(* IEC 61131-3 sources: plc-st-coding-agent/progress/evidence/f14_v13_self_20261113/jobs/custom_deepseek-v4pro (part 3) *)

(* ---- public-hard-05.patch_base_03.st ---- *)
FUNCTION_BLOCK MechanicalArmControl
VAR_INPUT
    ManualMode : BOOL;
    SingleStepMode : BOOL;
    SingleCycleMode : BOOL;
    ContinuousMode : BOOL;
    EmergencyStop : BOOL;
    Start : BOOL;
    DownButton : BOOL;
    UpButton : BOOL;
    LeftButton : BOOL;
    RightButton : BOOL;
    GripButton : BOOL;
    ReleaseButton : BOOL;
    DownLimitSwitch : BOOL;
    UpLimitSwitch : BOOL;
    LeftLimitSwitch : BOOL;
    RightLimitSwitch : BOOL;
    GripLimitSwitch : BOOL;
    ReleaseLimitSwitch : BOOL;
END_VAR
VAR_OUTPUT
    MoveDown : BOOL;
    MoveUp : BOOL;
    MoveLeft : BOOL;
    MoveRight : BOOL;
    ActivateGrip : BOOL;
    ActivateRelease : BOOL;
END_VAR
VAR
    local_startR : R_TRIG;
    tmp_first_scan : BOOL := TRUE;
    tmp_start_pulse : BOOL;
    tmp_not_estop : BOOL;
    tmp_ss_step : INT := 0;
    tmp_ss_busy : BOOL := FALSE;
    tmp_auto_running : BOOL := FALSE;
    tmp_auto_step : INT := 0;
    tmp_cmd_step : INT := 0;
    tmp_cmd_active : BOOL := FALSE;
    tmp_limit_reached : BOOL := FALSE;
END_VAR

(* ENGINEERING_CONTRACT
   Outputs MoveDown/Up/Left/Right/ActivateGrip/ActivateRelease:
   - Activate: manual while button=1, not at axis limit, and no opposite button (PUB001,PUB020); auto while current step active.
   - Retain: none latching; auto sequence state retained until completion/estop.
   - Reset: EmergencyStop=FALSE forces all outputs off and resets auto/single-step state (PUB005).
   - Same-scan: on limit true, previous output off; auto cycle can start next output in same scan (PUB003,PUB004).
   - Manual opposite-direction conflict inhibits both (PUB001 + shared rule).
   - Single-step Start edge only when not busy; ignored during running action (PUB002).
   - Single-cycle/continuous Start edge only when not running; continuous wraps at left completion (PUB003,PUB004).
   - Steps 0..7 = down, grip, up, right, down, release, up, left.
   - Grip/Release completion via GripLimitSwitch/ReleaseLimitSwitch (PUB001,PUB002).
   - Unspecified: mode change outside selected branch aborts/pauses per branch.
*)

(* CONTRACT_RULES [] *)

MoveDown := FALSE;
MoveUp := FALSE;
MoveLeft := FALSE;
MoveRight := FALSE;
ActivateGrip := FALSE;
ActivateRelease := FALSE;

tmp_not_estop := EmergencyStop; (* TRUE means no emergency stop triggered *)

local_startR(CLK := Start);
tmp_start_pulse := local_startR.Q AND NOT tmp_first_scan;
tmp_first_scan := FALSE;

tmp_cmd_active := FALSE;
tmp_cmd_step := 0;

IF NOT tmp_not_estop THEN
    tmp_ss_step := 0;
    tmp_ss_busy := FALSE;
    tmp_auto_running := FALSE;
    tmp_auto_step := 0;
    RETURN;
END_IF;

IF ManualMode THEN
    IF DownButton AND NOT UpButton AND NOT DownLimitSwitch THEN
        MoveDown := TRUE;
    END_IF;
    IF UpButton AND NOT DownButton AND NOT UpLimitSwitch THEN
        MoveUp := TRUE;
    END_IF;
    IF LeftButton AND NOT RightButton AND NOT LeftLimitSwitch THEN
        MoveLeft := TRUE;
    END_IF;
    IF RightButton AND NOT LeftButton AND NOT RightLimitSwitch THEN
        MoveRight := TRUE;
    END_IF;
    IF GripButton AND NOT ReleaseButton AND NOT GripLimitSwitch THEN
        ActivateGrip := TRUE;
    END_IF;
    IF ReleaseButton AND NOT GripButton AND NOT ReleaseLimitSwitch THEN
        ActivateRelease := TRUE;
    END_IF;

ELSIF SingleStepMode THEN
    IF tmp_start_pulse AND NOT tmp_ss_busy THEN
        tmp_ss_busy := TRUE;
    END_IF;

    IF tmp_ss_busy THEN
        tmp_limit_reached := FALSE;
        CASE tmp_ss_step OF
            0: tmp_limit_reached := DownLimitSwitch;
            1: tmp_limit_reached := GripLimitSwitch;
            2: tmp_limit_reached := UpLimitSwitch;
            3: tmp_limit_reached := RightLimitSwitch;
            4: tmp_limit_reached := DownLimitSwitch;
            5: tmp_limit_reached := ReleaseLimitSwitch;
            6: tmp_limit_reached := UpLimitSwitch;
            7: tmp_limit_reached := LeftLimitSwitch;
        END_CASE;

        IF tmp_limit_reached THEN
            tmp_ss_busy := FALSE;
            tmp_ss_step := tmp_ss_step + 1;
            IF tmp_ss_step > 7 THEN
                tmp_ss_step := 0;
            END_IF;
        ELSE
            tmp_cmd_step := tmp_ss_step;
            tmp_cmd_active := TRUE;
        END_IF;
    END_IF;

ELSIF SingleCycleMode OR ContinuousMode THEN
    IF tmp_start_pulse AND NOT tmp_auto_running THEN
        tmp_auto_running := TRUE;
        tmp_auto_step := 0;
    END_IF;

    IF tmp_auto_running THEN
        tmp_limit_reached := FALSE;
        CASE tmp_auto_step OF
            0: tmp_limit_reached := DownLimitSwitch;
            1: tmp_limit_reached := GripLimitSwitch;
            2: tmp_limit_reached := UpLimitSwitch;
            3: tmp_limit_reached := RightLimitSwitch;
            4: tmp_limit_reached := DownLimitSwitch;
            5: tmp_limit_reached := ReleaseLimitSwitch;
            6: tmp_limit_reached := UpLimitSwitch;
            7: tmp_limit_reached := LeftLimitSwitch;
        END_CASE;

        IF tmp_limit_reached THEN
            IF tmp_auto_step = 7 THEN
                IF ContinuousMode THEN
                    tmp_auto_step := 0; (* start next cycle *)
                ELSE
                    tmp_auto_running := FALSE;
                    tmp_auto_step := 0;
                END_IF;
            ELSE
                tmp_auto_step := tmp_auto_step + 1;
            END_IF;
        END_IF;

        IF tmp_auto_running THEN
            tmp_cmd_step := tmp_auto_step;
            tmp_cmd_active := TRUE;
        END_IF;
    END_IF;
END_IF;

IF tmp_cmd_active THEN
    CASE tmp_cmd_step OF
        0: MoveDown := TRUE;
        1: ActivateGrip := TRUE;
        2: MoveUp := TRUE;
        3: MoveRight := TRUE;
        4: MoveDown := TRUE;
        5: ActivateRelease := TRUE;
        6: MoveUp := TRUE;
        7: MoveLeft := TRUE;
    END_CASE;
END_IF;

END_FUNCTION_BLOCK

(* ---- public-hard-05.raw_candidate_01.st ---- *)
FUNCTION_BLOCK MechanicalArmControl
VAR_INPUT
    ManualMode : BOOL;
    SingleStepMode : BOOL;
    SingleCycleMode : BOOL;
    ContinuousMode : BOOL;
    EmergencyStop : BOOL;
    Start : BOOL;
    DownButton : BOOL;
    UpButton : BOOL;
    LeftButton : BOOL;
    RightButton : BOOL;
    GripButton : BOOL;
    ReleaseButton : BOOL;
    DownLimitSwitch : BOOL;
    UpLimitSwitch : BOOL;
    LeftLimitSwitch : BOOL;
    RightLimitSwitch : BOOL;
    GripLimitSwitch : BOOL;
    ReleaseLimitSwitch : BOOL;
END_VAR
VAR_OUTPUT
    MoveDown : BOOL;
    MoveUp : BOOL;
    MoveLeft : BOOL;
    MoveRight : BOOL;
    ActivateGrip : BOOL;
    ActivateRelease : BOOL;
END_VAR
VAR
    local_startR : R_TRIG;
    tmp_start_pulse : BOOL;
    tmp_not_estop : BOOL;
    tmp_ss_step : INT := 0;
    tmp_ss_busy : BOOL := FALSE;
    tmp_auto_running : BOOL := FALSE;
    tmp_auto_step : INT := 0;
    tmp_cmd_step : INT := 0;
    tmp_cmd_active : BOOL := FALSE;
    tmp_limit_reached : BOOL := FALSE;
END_VAR

(* ENGINEERING_CONTRACT
   Outputs MoveDown/Up/Left/Right/ActivateGrip/ActivateRelease:
   - Activate: manual while button=1, not at axis limit, and no opposite button (PUB001,PUB020); auto while current step active.
   - Retain: none latching; auto sequence state retained until completion/estop.
   - Reset: EmergencyStop=FALSE forces all outputs off and resets auto/single-step state (PUB005).
   - Same-scan: on limit true, previous output off; auto cycle can start next output in same scan (PUB003,PUB004).
   - Manual opposite-direction conflict inhibits both (PUB001 + shared rule).
   - Single-step Start edge only when not busy; ignored during running action (PUB002).
   - Single-cycle/continuous Start edge only when not running; continuous wraps at left completion (PUB003,PUB004).
   - Steps 0..7 = down, grip, up, right, down, release, up, left.
   - Grip/Release completion via GripLimitSwitch/ReleaseLimitSwitch (PUB001,PUB002).
   - Unspecified: mode change outside selected branch aborts/pauses per branch.
*)

(* CONTRACT_RULES [] *)

MoveDown := FALSE;
MoveUp := FALSE;
MoveLeft := FALSE;
MoveRight := FALSE;
ActivateGrip := FALSE;
ActivateRelease := FALSE;

tmp_not_estop := EmergencyStop; (* TRUE means no emergency stop triggered *)

local_startR(CLK := Start);
tmp_start_pulse := local_startR.Q;

tmp_cmd_active := FALSE;
tmp_cmd_step := 0;

IF NOT tmp_not_estop THEN
    tmp_ss_step := 0;
    tmp_ss_busy := FALSE;
    tmp_auto_running := FALSE;
    tmp_auto_step := 0;
    RETURN;
END_IF;

IF ManualMode THEN
    IF DownButton AND NOT UpButton AND NOT DownLimitSwitch THEN
        MoveDown := TRUE;
    END_IF;
    IF UpButton AND NOT DownButton AND NOT UpLimitSwitch THEN
        MoveUp := TRUE;
    END_IF;
    IF LeftButton AND NOT RightButton AND NOT LeftLimitSwitch THEN
        MoveLeft := TRUE;
    END_IF;
    IF RightButton AND NOT LeftButton AND NOT RightLimitSwitch THEN
        MoveRight := TRUE;
    END_IF;
    IF GripButton AND NOT ReleaseButton AND NOT GripLimitSwitch THEN
        ActivateGrip := TRUE;
    END_IF;
    IF ReleaseButton AND NOT GripButton AND NOT ReleaseLimitSwitch THEN
        ActivateRelease := TRUE;
    END_IF;

ELSIF SingleStepMode THEN
    IF tmp_start_pulse AND NOT tmp_ss_busy THEN
        tmp_ss_busy := TRUE;
    END_IF;

    IF tmp_ss_busy THEN
        tmp_limit_reached := FALSE;
        CASE tmp_ss_step OF
            0: tmp_limit_reached := DownLimitSwitch;
            1: tmp_limit_reached := GripLimitSwitch;
            2: tmp_limit_reached := UpLimitSwitch;
            3: tmp_limit_reached := RightLimitSwitch;
            4: tmp_limit_reached := DownLimitSwitch;
            5: tmp_limit_reached := ReleaseLimitSwitch;
            6: tmp_limit_reached := UpLimitSwitch;
            7: tmp_limit_reached := LeftLimitSwitch;
        END_CASE;

        IF tmp_limit_reached THEN
            tmp_ss_busy := FALSE;
            tmp_ss_step := tmp_ss_step + 1;
            IF tmp_ss_step > 7 THEN
                tmp_ss_step := 0;
            END_IF;
        ELSE
            tmp_cmd_step := tmp_ss_step;
            tmp_cmd_active := TRUE;
        END_IF;
    END_IF;

ELSIF SingleCycleMode OR ContinuousMode THEN
    IF tmp_start_pulse AND NOT tmp_auto_running THEN
        tmp_auto_running := TRUE;
        tmp_auto_step := 0;
    END_IF;

    IF tmp_auto_running THEN
        tmp_limit_reached := FALSE;
        CASE tmp_auto_step OF
            0: tmp_limit_reached := DownLimitSwitch;
            1: tmp_limit_reached := GripLimitSwitch;
            2: tmp_limit_reached := UpLimitSwitch;
            3: tmp_limit_reached := RightLimitSwitch;
            4: tmp_limit_reached := DownLimitSwitch;
            5: tmp_limit_reached := ReleaseLimitSwitch;
            6: tmp_limit_reached := UpLimitSwitch;
            7: tmp_limit_reached := LeftLimitSwitch;
        END_CASE;

        IF tmp_limit_reached THEN
            IF tmp_auto_step = 7 THEN
                IF ContinuousMode THEN
                    tmp_auto_step := 0; (* start next cycle *)
                ELSE
                    tmp_auto_running := FALSE;
                    tmp_auto_step := 0;
                END_IF;
            ELSE
                tmp_auto_step := tmp_auto_step + 1;
            END_IF;
        END_IF;

        IF tmp_auto_running THEN
            tmp_cmd_step := tmp_auto_step;
            tmp_cmd_active := TRUE;
        END_IF;
    END_IF;
END_IF;

IF tmp_cmd_active THEN
    CASE tmp_cmd_step OF
        0: MoveDown := TRUE;
        1: ActivateGrip := TRUE;
        2: MoveUp := TRUE;
        3: MoveRight := TRUE;
        4: MoveDown := TRUE;
        5: ActivateRelease := TRUE;
        6: MoveUp := TRUE;
        7: MoveLeft := TRUE;
    END_CASE;
END_IF;

END_FUNCTION_BLOCK

(* ---- public-hard-05.raw_candidate_02.st ---- *)
FUNCTION_BLOCK MechanicalArmControl
VAR_INPUT
    ManualMode : BOOL;
    SingleStepMode : BOOL;
    SingleCycleMode : BOOL;
    ContinuousMode : BOOL;
    EmergencyStop : BOOL;
    Start : BOOL;
    DownButton : BOOL;
    UpButton : BOOL;
    LeftButton : BOOL;
    RightButton : BOOL;
    GripButton : BOOL;
    ReleaseButton : BOOL;
    DownLimitSwitch : BOOL;
    UpLimitSwitch : BOOL;
    LeftLimitSwitch : BOOL;
    RightLimitSwitch : BOOL;
    GripLimitSwitch : BOOL;
    ReleaseLimitSwitch : BOOL;
END_VAR
VAR_OUTPUT
    MoveDown : BOOL;
    MoveUp : BOOL;
    MoveLeft : BOOL;
    MoveRight : BOOL;
    ActivateGrip : BOOL;
    ActivateRelease : BOOL;
END_VAR
VAR
    local_startR : R_TRIG;
    tmp_first_scan : BOOL := TRUE;
    tmp_start_pulse : BOOL;
    tmp_not_estop : BOOL;
    tmp_ss_step : INT := 0;
    tmp_ss_busy : BOOL := FALSE;
    tmp_auto_running : BOOL := FALSE;
    tmp_auto_step : INT := 0;
    tmp_cmd_step : INT := 0;
    tmp_cmd_active : BOOL := FALSE;
    tmp_limit_reached : BOOL := FALSE;
END_VAR

(* ENGINEERING_CONTRACT
   Outputs MoveDown/Up/Left/Right/ActivateGrip/ActivateRelease:
   - Activate: manual while button=1, not at axis limit, and no opposite button (PUB001,PUB020); auto while current step active.
   - Retain: none latching; auto sequence state retained until completion/estop.
   - Reset: EmergencyStop=FALSE forces all outputs off and resets auto/single-step state (PUB005).
   - Same-scan: on limit true, previous output off; auto cycle can start next output in same scan (PUB003,PUB004).
   - Manual opposite-direction conflict inhibits both (PUB001 + shared rule).
   - Single-step Start edge only when not busy; ignored during running action (PUB002).
   - Single-cycle/continuous Start edge only when not running; continuous wraps at left completion (PUB003,PUB004).
   - Steps 0..7 = down, grip, up, right, down, release, up, left.
   - Grip/Release completion via GripLimitSwitch/ReleaseLimitSwitch (PUB001,PUB002).
   - Unspecified: mode change outside selected branch aborts/pauses per branch.
*)

(* CONTRACT_RULES [] *)

MoveDown := FALSE;
MoveUp := FALSE;
MoveLeft := FALSE;
MoveRight := FALSE;
ActivateGrip := FALSE;
ActivateRelease := FALSE;

tmp_not_estop := EmergencyStop; (* TRUE means no emergency stop triggered *)

local_startR(CLK := Start);
tmp_start_pulse := local_startR.Q AND NOT tmp_first_scan;
tmp_first_scan := FALSE;

tmp_cmd_active := FALSE;
tmp_cmd_step := 0;

IF NOT tmp_not_estop THEN
    tmp_ss_step := 0;
    tmp_ss_busy := FALSE;
    tmp_auto_running := FALSE;
    tmp_auto_step := 0;
    RETURN;
END_IF;

IF ManualMode THEN
    IF DownButton AND NOT UpButton AND NOT DownLimitSwitch THEN
        MoveDown := TRUE;
    END_IF;
    IF UpButton AND NOT DownButton AND NOT UpLimitSwitch THEN
        MoveUp := TRUE;
    END_IF;
    IF LeftButton AND NOT RightButton AND NOT LeftLimitSwitch THEN
        MoveLeft := TRUE;
    END_IF;
    IF RightButton AND NOT LeftButton AND NOT RightLimitSwitch THEN
        MoveRight := TRUE;
    END_IF;
    IF GripButton AND NOT ReleaseButton AND NOT GripLimitSwitch THEN
        ActivateGrip := TRUE;
    END_IF;
    IF ReleaseButton AND NOT GripButton AND NOT ReleaseLimitSwitch THEN
        ActivateRelease := TRUE;
    END_IF;

ELSIF SingleStepMode THEN
    IF tmp_start_pulse AND NOT tmp_ss_busy THEN
        tmp_ss_busy := TRUE;
    END_IF;

    IF tmp_ss_busy THEN
        tmp_limit_reached := FALSE;
        CASE tmp_ss_step OF
            0: tmp_limit_reached := DownLimitSwitch;
            1: tmp_limit_reached := GripLimitSwitch;
            2: tmp_limit_reached := UpLimitSwitch;
            3: tmp_limit_reached := RightLimitSwitch;
            4: tmp_limit_reached := DownLimitSwitch;
            5: tmp_limit_reached := ReleaseLimitSwitch;
            6: tmp_limit_reached := UpLimitSwitch;
            7: tmp_limit_reached := LeftLimitSwitch;
        END_CASE;

        IF tmp_limit_reached THEN
            tmp_ss_busy := FALSE;
            tmp_ss_step := tmp_ss_step + 1;
            IF tmp_ss_step > 7 THEN
                tmp_ss_step := 0;
            END_IF;
        ELSE
            tmp_cmd_step := tmp_ss_step;
            tmp_cmd_active := TRUE;
        END_IF;
    END_IF;

ELSIF SingleCycleMode OR ContinuousMode THEN
    IF tmp_start_pulse AND NOT tmp_auto_running THEN
        tmp_auto_running := TRUE;
        tmp_auto_step := 0;
    END_IF;

    IF tmp_auto_running THEN
        tmp_limit_reached := FALSE;
        CASE tmp_auto_step OF
            0: tmp_limit_reached := DownLimitSwitch;
            1: tmp_limit_reached := GripLimitSwitch;
            2: tmp_limit_reached := UpLimitSwitch;
            3: tmp_limit_reached := RightLimitSwitch;
            4: tmp_limit_reached := DownLimitSwitch;
            5: tmp_limit_reached := ReleaseLimitSwitch;
            6: tmp_limit_reached := UpLimitSwitch;
            7: tmp_limit_reached := LeftLimitSwitch;
        END_CASE;

        IF tmp_limit_reached THEN
            IF tmp_auto_step = 7 THEN
                IF ContinuousMode THEN
                    tmp_auto_step := 0; (* start next cycle *)
                ELSE
                    tmp_auto_running := FALSE;
                    tmp_auto_step := 0;
                END_IF;
            ELSE
                tmp_auto_step := tmp_auto_step + 1;
            END_IF;
        END_IF;

        IF tmp_auto_running THEN
            tmp_cmd_step := tmp_auto_step;
            tmp_cmd_active := TRUE;
        END_IF;
    END_IF;
END_IF;

IF tmp_cmd_active THEN
    CASE tmp_cmd_step OF
        0: MoveDown := TRUE;
        1: ActivateGrip := TRUE;
        2: MoveUp := TRUE;
        3: MoveRight := TRUE;
        4: MoveDown := TRUE;
        5: ActivateRelease := TRUE;
        6: MoveUp := TRUE;
        7: MoveLeft := TRUE;
    END_CASE;
END_IF;

END_FUNCTION_BLOCK

(* ---- public-hard-05.raw_candidate_03.st ---- *)
FUNCTION_BLOCK MechanicalArmControl
VAR_INPUT
    ManualMode : BOOL;
    SingleStepMode : BOOL;
    SingleCycleMode : BOOL;
    ContinuousMode : BOOL;
    EmergencyStop : BOOL;
    Start : BOOL;
    DownButton : BOOL;
    UpButton : BOOL;
    LeftButton : BOOL;
    RightButton : BOOL;
    GripButton : BOOL;
    ReleaseButton : BOOL;
    DownLimitSwitch : BOOL;
    UpLimitSwitch : BOOL;
    LeftLimitSwitch : BOOL;
    RightLimitSwitch : BOOL;
    GripLimitSwitch : BOOL;
    ReleaseLimitSwitch : BOOL;
END_VAR
VAR_OUTPUT
    MoveDown : BOOL;
    MoveUp : BOOL;
    MoveLeft : BOOL;
    MoveRight : BOOL;
    ActivateGrip : BOOL;
    ActivateRelease : BOOL;
END_VAR
VAR
    local_startR : R_TRIG;
    tmp_start_pulse : BOOL;
    tmp_not_estop : BOOL;
    tmp_ss_step : INT := 0;
    tmp_ss_busy : BOOL := FALSE;
    tmp_auto_running : BOOL := FALSE;
    tmp_auto_step : INT := 0;
    tmp_cmd_step : INT := 0;
    tmp_cmd_active : BOOL := FALSE;
    tmp_limit_reached : BOOL := FALSE;
END_VAR

(* ENGINEERING_CONTRACT
   Outputs MoveDown/Up/Left/Right/ActivateGrip/ActivateRelease:
   - Activate: manual while button=1, not at axis limit, and no opposite button (PUB001,PUB020); auto while current step active.
   - Retain: none latching; auto sequence state retained until completion/estop.
   - Reset: EmergencyStop=FALSE forces all outputs off and resets auto/single-step state (PUB005).
   - Same-scan: on limit true, previous output off; auto cycle can start next output in same scan (PUB003,PUB004).
   - Manual opposite-direction conflict inhibits both (PUB001 + shared rule).
   - Single-step Start edge only when not busy; ignored during running action (PUB002).
   - Single-cycle/continuous Start edge only when not running; continuous wraps at left completion (PUB003,PUB004).
   - Steps 0..7 = down, grip, up, right, down, release, up, left.
   - Grip/Release completion via GripLimitSwitch/ReleaseLimitSwitch (PUB001,PUB002).
   - Unspecified: mode change outside selected branch aborts/pauses per branch.
*)

(* CONTRACT_RULES [] *)

MoveDown := FALSE;
MoveUp := FALSE;
MoveLeft := FALSE;
MoveRight := FALSE;
ActivateGrip := FALSE;
ActivateRelease := FALSE;

tmp_not_estop := EmergencyStop; (* TRUE means no emergency stop triggered *)

local_startR(CLK := Start);
tmp_start_pulse := local_startR.Q;

tmp_cmd_active := FALSE;
tmp_cmd_step := 0;

IF NOT tmp_not_estop THEN
    tmp_ss_step := 0;
    tmp_ss_busy := FALSE;
    tmp_auto_running := FALSE;
    tmp_auto_step := 0;
    RETURN;
END_IF;

IF ManualMode THEN
    IF DownButton AND NOT UpButton AND NOT DownLimitSwitch THEN
        MoveDown := TRUE;
    END_IF;
    IF UpButton AND NOT DownButton AND NOT UpLimitSwitch THEN
        MoveUp := TRUE;
    END_IF;
    IF LeftButton AND NOT RightButton AND NOT LeftLimitSwitch THEN
        MoveLeft := TRUE;
    END_IF;
    IF RightButton AND NOT LeftButton AND NOT RightLimitSwitch THEN
        MoveRight := TRUE;
    END_IF;
    IF GripButton AND NOT ReleaseButton AND NOT GripLimitSwitch THEN
        ActivateGrip := TRUE;
    END_IF;
    IF ReleaseButton AND NOT GripButton AND NOT ReleaseLimitSwitch THEN
        ActivateRelease := TRUE;
    END_IF;

ELSIF SingleStepMode THEN
    IF tmp_start_pulse AND NOT tmp_ss_busy THEN
        tmp_ss_busy := TRUE;
    END_IF;

    IF tmp_ss_busy THEN
        tmp_limit_reached := FALSE;
        CASE tmp_ss_step OF
            0: tmp_limit_reached := DownLimitSwitch;
            1: tmp_limit_reached := GripLimitSwitch;
            2: tmp_limit_reached := UpLimitSwitch;
            3: tmp_limit_reached := RightLimitSwitch;
            4: tmp_limit_reached := DownLimitSwitch;
            5: tmp_limit_reached := ReleaseLimitSwitch;
            6: tmp_limit_reached := UpLimitSwitch;
            7: tmp_limit_reached := LeftLimitSwitch;
        END_CASE;

        IF tmp_limit_reached THEN
            tmp_ss_busy := FALSE;
            tmp_ss_step := tmp_ss_step + 1;
            IF tmp_ss_step > 7 THEN
                tmp_ss_step := 0;
            END_IF;
        ELSE
            tmp_cmd_step := tmp_ss_step;
            tmp_cmd_active := TRUE;
        END_IF;
    END_IF;

ELSIF SingleCycleMode OR ContinuousMode THEN
    IF tmp_start_pulse AND NOT tmp_auto_running THEN
        tmp_auto_running := TRUE;
        tmp_auto_step := 0;
    END_IF;

    IF tmp_auto_running THEN
        tmp_limit_reached := FALSE;
        CASE tmp_auto_step OF
            0: tmp_limit_reached := DownLimitSwitch;
            1: tmp_limit_reached := GripLimitSwitch;
            2: tmp_limit_reached := UpLimitSwitch;
            3: tmp_limit_reached := RightLimitSwitch;
            4: tmp_limit_reached := DownLimitSwitch;
            5: tmp_limit_reached := ReleaseLimitSwitch;
            6: tmp_limit_reached := UpLimitSwitch;
            7: tmp_limit_reached := LeftLimitSwitch;
        END_CASE;

        IF tmp_limit_reached THEN
            IF tmp_auto_step = 7 THEN
                IF ContinuousMode THEN
                    tmp_auto_step := 0; (* start next cycle *)
                ELSE
                    tmp_auto_running := FALSE;
                    tmp_auto_step := 0;
                END_IF;
            ELSE
                tmp_auto_step := tmp_auto_step + 1;
            END_IF;
        END_IF;

        IF tmp_auto_running THEN
            tmp_cmd_step := tmp_auto_step;
            tmp_cmd_active := TRUE;
        END_IF;
    END_IF;
END_IF;

IF tmp_cmd_active THEN
    CASE tmp_cmd_step OF
        0: MoveDown := TRUE;
        1: ActivateGrip := TRUE;
        2: MoveUp := TRUE;
        3: MoveRight := TRUE;
        4: MoveDown := TRUE;
        5: ActivateRelease := TRUE;
        6: MoveUp := TRUE;
        7: MoveLeft := TRUE;
    END_CASE;
END_IF;

END_FUNCTION_BLOCK

(* ---- public-hard-06.candidate_01.st ---- *)
FUNCTION_BLOCK ProductionControl
VAR_INPUT
    Mode : BOOL;
    ForwardButton : BOOL;
    ReverseButton : BOOL;
    SensorFeed : BOOL;
    SensorWash : BOOL;
    SensorWeight : BOOL;
    SensorFiring : BOOL;
    SensorOutput : BOOL;
    washComplete : BOOL;
    weightComplete : BOOL;
    weight : REAL;
    firingComplete : BOOL;
END_VAR
VAR_OUTPUT
    MotorForward : BOOL;
    MotorReverse : BOOL;
    kick : BOOL;
    CompletionLight : BOOL;
    firingTemp : REAL;
END_VAR
VAR
    AutoStep : INT := 0;
    AutoInit : BOOL := FALSE;
    lastFiringTemp : REAL := 0.0;
    rtWash : R_TRIG;
    rtWeight : R_TRIG;
    rtFiring : R_TRIG;
    washEdge : BOOL;
    weightEdge : BOOL;
    firingEdge : BOOL;
    tmp_unqualified : BOOL;
END_VAR

(*
ENGINEERING_CONTRACT
MotorForward: auto active in states 10/30/50/70; manual = ForwardButton AND NOT ReverseButton.
MotorReverse: manual only, interlocked with ForwardButton; both false if both buttons true.
kick: pulse on rising weightComplete when weight < 100 or weight > 200 (unqualified).
CompletionLight: combinational = SensorOutput while Mode=TRUE; off in manual.
firingTemp: stored on qualified weightComplete; formula 500 + (weight-100)*0.5, retained otherwise.
Units: weight REAL in same unit as thresholds; firingTemp REAL degrees; boundaries inclusive 100..200.
*)
(* CONTRACT_RULES [] *)

rtWash(CLK := washComplete);
rtWeight(CLK := weightComplete);
rtFiring(CLK := firingComplete);
washEdge := rtWash.Q;
weightEdge := rtWeight.Q;
firingEdge := rtFiring.Q;

IF NOT AutoInit THEN
    AutoInit := TRUE;
    IF SensorOutput THEN
        AutoStep := 80;
    ELSIF SensorFiring THEN
        AutoStep := 60;
    ELSIF SensorWeight THEN
        AutoStep := 40;
    ELSIF SensorWash THEN
        AutoStep := 20;
    ELSIF SensorFeed THEN
        AutoStep := 10;
    ELSE
        AutoStep := 0;
    END_IF;
END_IF;

IF NOT Mode THEN
    MotorForward := ForwardButton AND (NOT ReverseButton);
    MotorReverse := ReverseButton AND (NOT ForwardButton);
    kick := FALSE;
    CompletionLight := FALSE;
    firingTemp := lastFiringTemp;
    RETURN;
END_IF;

MotorForward := FALSE;
MotorReverse := FALSE;
kick := FALSE;
CompletionLight := FALSE;

CASE AutoStep OF
    0:
        IF SensorFeed THEN
            AutoStep := 10;
        END_IF;

    10:
        IF SensorWash THEN
            AutoStep := 20;
        END_IF;

    20:
        IF washEdge THEN
            AutoStep := 30;
        END_IF;

    30:
        IF SensorWeight THEN
            AutoStep := 40;
        END_IF;

    40:
        IF weightEdge THEN
            tmp_unqualified := (weight < 100.0) OR (weight > 200.0);
            IF tmp_unqualified THEN
                kick := TRUE;
                AutoStep := 0;
            ELSE
                lastFiringTemp := 500.0 + (weight - 100.0) * 0.5;
                AutoStep := 50;
            END_IF;
        END_IF;

    50:
        IF SensorFiring THEN
            AutoStep := 60;
        END_IF;

    60:
        IF firingEdge THEN
            AutoStep := 70;
        END_IF;

    70:
        IF SensorOutput THEN
            AutoStep := 80;
        END_IF;

    80:
        ;
END_CASE;

MotorForward := (AutoStep = 10) OR (AutoStep = 30) OR (AutoStep = 50) OR (AutoStep = 70);
MotorReverse := FALSE;
CompletionLight := SensorOutput;
firingTemp := lastFiringTemp;
END_FUNCTION_BLOCK

(* ---- public-hard-06.candidate_02.st ---- *)
FUNCTION_BLOCK ProductionControl
VAR_INPUT
    Mode : BOOL;
    ForwardButton : BOOL;
    ReverseButton : BOOL;
    SensorFeed : BOOL;
    SensorWash : BOOL;
    SensorWeight : BOOL;
    SensorFiring : BOOL;
    SensorOutput : BOOL;
    washComplete : BOOL;
    weightComplete : BOOL;
    weight : REAL;
    firingComplete : BOOL;
END_VAR
VAR_OUTPUT
    MotorForward : BOOL;
    MotorReverse : BOOL;
    kick : BOOL;
    CompletionLight : BOOL;
    firingTemp : REAL;
END_VAR
VAR
    AutoStep : INT := 0;
    AutoInit : BOOL := FALSE;
    lastFiringTemp : REAL := 0.0;
    rtWash : R_TRIG;
    rtWeight : R_TRIG;
    rtFiring : R_TRIG;
    washEdge : BOOL;
    weightEdge : BOOL;
    firingEdge : BOOL;
    tmp_unqualified : BOOL;
END_VAR

(*
ENGINEERING_CONTRACT
MotorForward: auto active in states 10/30/50/70; manual = ForwardButton AND NOT ReverseButton.
MotorReverse: manual only, interlocked with ForwardButton; both false if both buttons true.
kick: pulse on rising weightComplete when weight < 100 or weight > 200 (unqualified).
CompletionLight: combinational = SensorOutput while Mode=TRUE; off in manual.
firingTemp: stored on qualified weightComplete; formula 500 + (weight-100)*0.5, retained otherwise.
Units: weight REAL in same unit as thresholds; firingTemp REAL degrees; boundaries inclusive 100..200.
*)
(* CONTRACT_RULES [] *)

rtWash(CLK := washComplete);
rtWeight(CLK := weightComplete);
rtFiring(CLK := firingComplete);
washEdge := rtWash.Q;
weightEdge := rtWeight.Q;
firingEdge := rtFiring.Q;

IF NOT AutoInit THEN
    AutoInit := TRUE;
    IF SensorOutput THEN
        AutoStep := 80;
    ELSIF SensorFiring THEN
        AutoStep := 60;
    ELSIF SensorWeight THEN
        AutoStep := 40;
    ELSIF SensorWash THEN
        AutoStep := 20;
    ELSIF SensorFeed THEN
        AutoStep := 10;
    ELSE
        AutoStep := 0;
    END_IF;
END_IF;

IF NOT Mode THEN
    MotorForward := ForwardButton AND (NOT ReverseButton);
    MotorReverse := ReverseButton AND (NOT ForwardButton);
    kick := FALSE;
    CompletionLight := FALSE;
    firingTemp := lastFiringTemp;
    RETURN;
END_IF;

MotorForward := FALSE;
MotorReverse := FALSE;
kick := FALSE;
CompletionLight := FALSE;

CASE AutoStep OF
    0:
        IF SensorFeed THEN
            AutoStep := 10;
        END_IF;

    10:
        IF SensorWash THEN
            AutoStep := 20;
        END_IF;

    20:
        IF washEdge THEN
            AutoStep := 30;
        END_IF;

    30:
        IF SensorWeight THEN
            AutoStep := 40;
        END_IF;

    40:
        IF weightEdge THEN
            tmp_unqualified := (weight < 100.0) OR (weight > 200.0);
            IF tmp_unqualified THEN
                kick := TRUE;
                AutoStep := 0;
            ELSE
                lastFiringTemp := 500.0 + (weight - 100.0) * 0.5;
                AutoStep := 50;
            END_IF;
        END_IF;

    50:
        IF SensorFiring THEN
            AutoStep := 60;
        END_IF;

    60:
        IF firingEdge THEN
            AutoStep := 70;
        END_IF;

    70:
        IF SensorOutput THEN
            AutoStep := 80;
        END_IF;

    80:
        IF NOT SensorOutput THEN
            AutoStep := 0;
        END_IF;
END_CASE;

MotorForward := (AutoStep = 10) OR (AutoStep = 30) OR (AutoStep = 50) OR (AutoStep = 70);
MotorReverse := FALSE;
CompletionLight := SensorOutput;
firingTemp := lastFiringTemp;
END_FUNCTION_BLOCK

(* ---- public-hard-06.candidate_03.st ---- *)
FUNCTION_BLOCK ProductionControl
VAR_INPUT
    Mode : BOOL;
    ForwardButton : BOOL;
    ReverseButton : BOOL;
    SensorFeed : BOOL;
    SensorWash : BOOL;
    SensorWeight : BOOL;
    SensorFiring : BOOL;
    SensorOutput : BOOL;
    washComplete : BOOL;
    weightComplete : BOOL;
    weight : REAL;
    firingComplete : BOOL;
END_VAR
VAR_OUTPUT
    MotorForward : BOOL;
    MotorReverse : BOOL;
    kick : BOOL;
    CompletionLight : BOOL;
    firingTemp : REAL;
END_VAR
VAR
    AutoStep : INT := 0;
    AutoInit : BOOL := FALSE;
    lastFiringTemp : REAL := 0.0;
    rtWash : R_TRIG;
    rtWeight : R_TRIG;
    rtFiring : R_TRIG;
    washEdge : BOOL;
    weightEdge : BOOL;
    firingEdge : BOOL;
    rtMode : R_TRIG;
    ModeRise : BOOL;
    tmp_unqualified : BOOL;
END_VAR

(*
ENGINEERING_CONTRACT
MotorForward: auto active in states 10/30/50/70; manual = ForwardButton AND NOT ReverseButton.
MotorReverse: manual only, interlocked with ForwardButton; both false if both buttons true.
kick: pulse on rising weightComplete when weight < 100 or weight > 200 (unqualified).
CompletionLight: combinational = SensorOutput while Mode=TRUE; off in manual.
firingTemp: stored on qualified weightComplete; formula 500 + (weight-100)*0.5, retained otherwise.
Units: weight REAL in same unit as thresholds; firingTemp REAL degrees; boundaries inclusive 100..200.
*)
(* CONTRACT_RULES [] *)

rtMode(CLK := Mode);
ModeRise := rtMode.Q;
rtWash(CLK := washComplete);
rtWeight(CLK := weightComplete);
rtFiring(CLK := firingComplete);
washEdge := rtWash.Q;
weightEdge := rtWeight.Q;
firingEdge := rtFiring.Q;

IF (NOT AutoInit) OR ModeRise THEN
    AutoInit := TRUE;
    IF SensorOutput THEN
        AutoStep := 80;
    ELSIF SensorFiring THEN
        AutoStep := 60;
    ELSIF SensorWeight THEN
        AutoStep := 40;
    ELSIF SensorWash THEN
        AutoStep := 20;
    ELSIF SensorFeed THEN
        AutoStep := 10;
    ELSE
        AutoStep := 0;
    END_IF;
END_IF;

IF NOT Mode THEN
    MotorForward := ForwardButton AND (NOT ReverseButton);
    MotorReverse := ReverseButton AND (NOT ForwardButton);
    kick := FALSE;
    CompletionLight := FALSE;
    firingTemp := lastFiringTemp;
    RETURN;
END_IF;

MotorForward := FALSE;
MotorReverse := FALSE;
kick := FALSE;
CompletionLight := FALSE;

CASE AutoStep OF
    0:
        IF SensorFeed THEN
            AutoStep := 10;
        END_IF;

    10:
        IF SensorWash THEN
            AutoStep := 20;
        END_IF;

    20:
        IF washEdge THEN
            AutoStep := 30;
        END_IF;

    30:
        IF SensorWeight THEN
            AutoStep := 40;
        END_IF;

    40:
        IF weightEdge THEN
            tmp_unqualified := (weight < 100.0) OR (weight > 200.0);
            IF tmp_unqualified THEN
                kick := TRUE;
                AutoStep := 0;
            ELSE
                lastFiringTemp := 500.0 + (weight - 100.0) * 0.5;
                AutoStep := 50;
            END_IF;
        END_IF;

    50:
        IF SensorFiring THEN
            AutoStep := 60;
        END_IF;

    60:
        IF firingEdge THEN
            AutoStep := 70;
        END_IF;

    70:
        IF SensorOutput THEN
            AutoStep := 80;
        END_IF;

    80:
        IF NOT SensorOutput THEN
            AutoStep := 0;
        END_IF;
END_CASE;

MotorForward := (AutoStep = 10) OR (AutoStep = 30) OR (AutoStep = 50) OR (AutoStep = 70);
MotorReverse := FALSE;
CompletionLight := SensorOutput;
firingTemp := lastFiringTemp;
END_FUNCTION_BLOCK

(* ---- public-hard-06.candidate_04.st ---- *)
FUNCTION_BLOCK ProductionControl
VAR_INPUT
    Mode : BOOL;
    ForwardButton : BOOL;
    ReverseButton : BOOL;
    SensorFeed : BOOL;
    SensorWash : BOOL;
    SensorWeight : BOOL;
    SensorFiring : BOOL;
    SensorOutput : BOOL;
    washComplete : BOOL;
    weightComplete : BOOL;
    weight : REAL;
    firingComplete : BOOL;
END_VAR
VAR_OUTPUT
    MotorForward : BOOL;
    MotorReverse : BOOL;
    kick : BOOL;
    CompletionLight : BOOL;
    firingTemp : REAL;
END_VAR
VAR
    AutoStep : INT := 0;
    AutoInit : BOOL := FALSE;
    lastFiringTemp : REAL := 0.0;
    rtWash : R_TRIG;
    rtWeight : R_TRIG;
    rtFiring : R_TRIG;
    washEdge : BOOL;
    weightEdge : BOOL;
    firingEdge : BOOL;
    rtMode : R_TRIG;
    ModeRise : BOOL;
    tmp_unqualified : BOOL;
END_VAR

(*
ENGINEERING_CONTRACT
MotorForward: auto active in states 10/30/50/70; manual = ForwardButton AND NOT ReverseButton.
MotorReverse: manual only, interlocked with ForwardButton; both false if both buttons true.
kick: pulse on rising weightComplete when weight < 100 or weight > 200 (unqualified).
CompletionLight: combinational = SensorOutput while Mode=TRUE; off in manual.
firingTemp: stored on qualified weightComplete; formula 500 + (weight-100)*0.5, retained otherwise.
Units: weight REAL in same unit as thresholds; firingTemp REAL degrees; boundaries inclusive 100..200.
*)
(* CONTRACT_RULES [] *)

rtMode(CLK := Mode);
ModeRise := rtMode.Q;
rtWash(CLK := washComplete);
rtWeight(CLK := weightComplete);
rtFiring(CLK := firingComplete);
washEdge := rtWash.Q;
weightEdge := rtWeight.Q;
firingEdge := rtFiring.Q;

IF (NOT AutoInit) OR ModeRise THEN
    AutoInit := TRUE;
    IF SensorOutput THEN
        AutoStep := 80;
    ELSIF SensorFiring THEN
        AutoStep := 60;
    ELSIF SensorWeight THEN
        AutoStep := 40;
    ELSIF SensorWash THEN
        AutoStep := 20;
    ELSIF SensorFeed THEN
        AutoStep := 10;
    ELSE
        AutoStep := 0;
    END_IF;
END_IF;

IF NOT Mode THEN
    MotorForward := ForwardButton AND (NOT ReverseButton);
    MotorReverse := ReverseButton AND (NOT ForwardButton);
    kick := FALSE;
    CompletionLight := FALSE;
    firingTemp := lastFiringTemp;
    RETURN;
END_IF;

MotorForward := FALSE;
MotorReverse := FALSE;
kick := FALSE;
CompletionLight := FALSE;

CASE AutoStep OF
    0:
        IF SensorFeed THEN
            AutoStep := 10;
        END_IF;

    10:
        IF SensorWash THEN
            AutoStep := 20;
        END_IF;

    20:
        IF washComplete THEN
            AutoStep := 30;
        END_IF;

    30:
        IF SensorWeight THEN
            AutoStep := 40;
        END_IF;

    40:
        IF weightComplete THEN
            tmp_unqualified := (weight < 100.0) OR (weight > 200.0);
            IF tmp_unqualified THEN
                kick := TRUE;
                AutoStep := 0;
            ELSE
                lastFiringTemp := 500.0 + (weight - 100.0) * 0.5;
                AutoStep := 50;
            END_IF;
        END_IF;

    50:
        IF SensorFiring THEN
            AutoStep := 60;
        END_IF;

    60:
        IF firingComplete THEN
            AutoStep := 70;
        END_IF;

    70:
        IF SensorOutput THEN
            AutoStep := 80;
        END_IF;

    80:
        IF NOT SensorOutput THEN
            AutoStep := 0;
        END_IF;
END_CASE;

MotorForward := (AutoStep = 10) OR (AutoStep = 30) OR (AutoStep = 50) OR (AutoStep = 70);
MotorReverse := FALSE;
CompletionLight := SensorOutput;
firingTemp := lastFiringTemp;
END_FUNCTION_BLOCK

(* ---- public-hard-06.patch_base_02.st ---- *)
FUNCTION_BLOCK ProductionControl
VAR_INPUT
    Mode : BOOL;
    ForwardButton : BOOL;
    ReverseButton : BOOL;
    SensorFeed : BOOL;
    SensorWash : BOOL;
    SensorWeight : BOOL;
    SensorFiring : BOOL;
    SensorOutput : BOOL;
    washComplete : BOOL;
    weightComplete : BOOL;
    weight : REAL;
    firingComplete : BOOL;
END_VAR
VAR_OUTPUT
    MotorForward : BOOL;
    MotorReverse : BOOL;
    kick : BOOL;
    CompletionLight : BOOL;
    firingTemp : REAL;
END_VAR
VAR
    AutoStep : INT := 0;
    AutoInit : BOOL := FALSE;
    lastFiringTemp : REAL := 0.0;
    rtWash : R_TRIG;
    rtWeight : R_TRIG;
    rtFiring : R_TRIG;
    washEdge : BOOL;
    weightEdge : BOOL;
    firingEdge : BOOL;
    tmp_unqualified : BOOL;
END_VAR

(*
ENGINEERING_CONTRACT
MotorForward: auto active in states 10/30/50/70; manual = ForwardButton AND NOT ReverseButton.
MotorReverse: manual only, interlocked with ForwardButton; both false if both buttons true.
kick: pulse on rising weightComplete when weight < 100 or weight > 200 (unqualified).
CompletionLight: combinational = SensorOutput while Mode=TRUE; off in manual.
firingTemp: stored on qualified weightComplete; formula 500 + (weight-100)*0.5, retained otherwise.
Units: weight REAL in same unit as thresholds; firingTemp REAL degrees; boundaries inclusive 100..200.
*)
(* CONTRACT_RULES [] *)

rtWash(CLK := washComplete);
rtWeight(CLK := weightComplete);
rtFiring(CLK := firingComplete);
washEdge := rtWash.Q;
weightEdge := rtWeight.Q;
firingEdge := rtFiring.Q;

IF NOT AutoInit THEN
    AutoInit := TRUE;
    IF SensorOutput THEN
        AutoStep := 80;
    ELSIF SensorFiring THEN
        AutoStep := 60;
    ELSIF SensorWeight THEN
        AutoStep := 40;
    ELSIF SensorWash THEN
        AutoStep := 20;
    ELSIF SensorFeed THEN
        AutoStep := 10;
    ELSE
        AutoStep := 0;
    END_IF;
END_IF;

IF NOT Mode THEN
    MotorForward := ForwardButton AND (NOT ReverseButton);
    MotorReverse := ReverseButton AND (NOT ForwardButton);
    kick := FALSE;
    CompletionLight := FALSE;
    firingTemp := lastFiringTemp;
    RETURN;
END_IF;

MotorForward := FALSE;
MotorReverse := FALSE;
kick := FALSE;
CompletionLight := FALSE;

CASE AutoStep OF
    0:
        IF SensorFeed THEN
            AutoStep := 10;
        END_IF;

    10:
        IF SensorWash THEN
            AutoStep := 20;
        END_IF;

    20:
        IF washEdge THEN
            AutoStep := 30;
        END_IF;

    30:
        IF SensorWeight THEN
            AutoStep := 40;
        END_IF;

    40:
        IF weightEdge THEN
            tmp_unqualified := (weight < 100.0) OR (weight > 200.0);
            IF tmp_unqualified THEN
                kick := TRUE;
                AutoStep := 0;
            ELSE
                lastFiringTemp := 500.0 + (weight - 100.0) * 0.5;
                AutoStep := 50;
            END_IF;
        END_IF;

    50:
        IF SensorFiring THEN
            AutoStep := 60;
        END_IF;

    60:
        IF firingEdge THEN
            AutoStep := 70;
        END_IF;

    70:
        IF SensorOutput THEN
            AutoStep := 80;
        END_IF;

    80:
        ;
END_CASE;

MotorForward := (AutoStep = 10) OR (AutoStep = 30) OR (AutoStep = 50) OR (AutoStep = 70);
MotorReverse := FALSE;
CompletionLight := SensorOutput;
firingTemp := lastFiringTemp;
END_FUNCTION_BLOCK

(* ---- public-hard-06.patch_base_03.st ---- *)
FUNCTION_BLOCK ProductionControl
VAR_INPUT
    Mode : BOOL;
    ForwardButton : BOOL;
    ReverseButton : BOOL;
    SensorFeed : BOOL;
    SensorWash : BOOL;
    SensorWeight : BOOL;
    SensorFiring : BOOL;
    SensorOutput : BOOL;
    washComplete : BOOL;
    weightComplete : BOOL;
    weight : REAL;
    firingComplete : BOOL;
END_VAR
VAR_OUTPUT
    MotorForward : BOOL;
    MotorReverse : BOOL;
    kick : BOOL;
    CompletionLight : BOOL;
    firingTemp : REAL;
END_VAR
VAR
    AutoStep : INT := 0;
    AutoInit : BOOL := FALSE;
    lastFiringTemp : REAL := 0.0;
    rtWash : R_TRIG;
    rtWeight : R_TRIG;
    rtFiring : R_TRIG;
    washEdge : BOOL;
    weightEdge : BOOL;
    firingEdge : BOOL;
    tmp_unqualified : BOOL;
END_VAR

(*
ENGINEERING_CONTRACT
MotorForward: auto active in states 10/30/50/70; manual = ForwardButton AND NOT ReverseButton.
MotorReverse: manual only, interlocked with ForwardButton; both false if both buttons true.
kick: pulse on rising weightComplete when weight < 100 or weight > 200 (unqualified).
CompletionLight: combinational = SensorOutput while Mode=TRUE; off in manual.
firingTemp: stored on qualified weightComplete; formula 500 + (weight-100)*0.5, retained otherwise.
Units: weight REAL in same unit as thresholds; firingTemp REAL degrees; boundaries inclusive 100..200.
*)
(* CONTRACT_RULES [] *)

rtWash(CLK := washComplete);
rtWeight(CLK := weightComplete);
rtFiring(CLK := firingComplete);
washEdge := rtWash.Q;
weightEdge := rtWeight.Q;
firingEdge := rtFiring.Q;

IF NOT AutoInit THEN
    AutoInit := TRUE;
    IF SensorOutput THEN
        AutoStep := 80;
    ELSIF SensorFiring THEN
        AutoStep := 60;
    ELSIF SensorWeight THEN
        AutoStep := 40;
    ELSIF SensorWash THEN
        AutoStep := 20;
    ELSIF SensorFeed THEN
        AutoStep := 10;
    ELSE
        AutoStep := 0;
    END_IF;
END_IF;

IF NOT Mode THEN
    MotorForward := ForwardButton AND (NOT ReverseButton);
    MotorReverse := ReverseButton AND (NOT ForwardButton);
    kick := FALSE;
    CompletionLight := FALSE;
    firingTemp := lastFiringTemp;
    RETURN;
END_IF;

MotorForward := FALSE;
MotorReverse := FALSE;
kick := FALSE;
CompletionLight := FALSE;

CASE AutoStep OF
    0:
        IF SensorFeed THEN
            AutoStep := 10;
        END_IF;

    10:
        IF SensorWash THEN
            AutoStep := 20;
        END_IF;

    20:
        IF washEdge THEN
            AutoStep := 30;
        END_IF;

    30:
        IF SensorWeight THEN
            AutoStep := 40;
        END_IF;

    40:
        IF weightEdge THEN
            tmp_unqualified := (weight < 100.0) OR (weight > 200.0);
            IF tmp_unqualified THEN
                kick := TRUE;
                AutoStep := 0;
            ELSE
                lastFiringTemp := 500.0 + (weight - 100.0) * 0.5;
                AutoStep := 50;
            END_IF;
        END_IF;

    50:
        IF SensorFiring THEN
            AutoStep := 60;
        END_IF;

    60:
        IF firingEdge THEN
            AutoStep := 70;
        END_IF;

    70:
        IF SensorOutput THEN
            AutoStep := 80;
        END_IF;

    80:
        IF NOT SensorOutput THEN
            AutoStep := 0;
        END_IF;
END_CASE;

MotorForward := (AutoStep = 10) OR (AutoStep = 30) OR (AutoStep = 50) OR (AutoStep = 70);
MotorReverse := FALSE;
CompletionLight := SensorOutput;
firingTemp := lastFiringTemp;
END_FUNCTION_BLOCK

(* ---- public-hard-06.patch_base_04.st ---- *)
FUNCTION_BLOCK ProductionControl
VAR_INPUT
    Mode : BOOL;
    ForwardButton : BOOL;
    ReverseButton : BOOL;
    SensorFeed : BOOL;
    SensorWash : BOOL;
    SensorWeight : BOOL;
    SensorFiring : BOOL;
    SensorOutput : BOOL;
    washComplete : BOOL;
    weightComplete : BOOL;
    weight : REAL;
    firingComplete : BOOL;
END_VAR
VAR_OUTPUT
    MotorForward : BOOL;
    MotorReverse : BOOL;
    kick : BOOL;
    CompletionLight : BOOL;
    firingTemp : REAL;
END_VAR
VAR
    AutoStep : INT := 0;
    AutoInit : BOOL := FALSE;
    lastFiringTemp : REAL := 0.0;
    rtWash : R_TRIG;
    rtWeight : R_TRIG;
    rtFiring : R_TRIG;
    washEdge : BOOL;
    weightEdge : BOOL;
    firingEdge : BOOL;
    rtMode : R_TRIG;
    ModeRise : BOOL;
    tmp_unqualified : BOOL;
END_VAR

(*
ENGINEERING_CONTRACT
MotorForward: auto active in states 10/30/50/70; manual = ForwardButton AND NOT ReverseButton.
MotorReverse: manual only, interlocked with ForwardButton; both false if both buttons true.
kick: pulse on rising weightComplete when weight < 100 or weight > 200 (unqualified).
CompletionLight: combinational = SensorOutput while Mode=TRUE; off in manual.
firingTemp: stored on qualified weightComplete; formula 500 + (weight-100)*0.5, retained otherwise.
Units: weight REAL in same unit as thresholds; firingTemp REAL degrees; boundaries inclusive 100..200.
*)
(* CONTRACT_RULES [] *)

rtMode(CLK := Mode);
ModeRise := rtMode.Q;
rtWash(CLK := washComplete);
rtWeight(CLK := weightComplete);
rtFiring(CLK := firingComplete);
washEdge := rtWash.Q;
weightEdge := rtWeight.Q;
firingEdge := rtFiring.Q;

IF (NOT AutoInit) OR ModeRise THEN
    AutoInit := TRUE;
    IF SensorOutput THEN
        AutoStep := 80;
    ELSIF SensorFiring THEN
        AutoStep := 60;
    ELSIF SensorWeight THEN
        AutoStep := 40;
    ELSIF SensorWash THEN
        AutoStep := 20;
    ELSIF SensorFeed THEN
        AutoStep := 10;
    ELSE
        AutoStep := 0;
    END_IF;
END_IF;

IF NOT Mode THEN
    MotorForward := ForwardButton AND (NOT ReverseButton);
    MotorReverse := ReverseButton AND (NOT ForwardButton);
    kick := FALSE;
    CompletionLight := FALSE;
    firingTemp := lastFiringTemp;
    RETURN;
END_IF;

MotorForward := FALSE;
MotorReverse := FALSE;
kick := FALSE;
CompletionLight := FALSE;

CASE AutoStep OF
    0:
        IF SensorFeed THEN
            AutoStep := 10;
        END_IF;

    10:
        IF SensorWash THEN
            AutoStep := 20;
        END_IF;

    20:
        IF washEdge THEN
            AutoStep := 30;
        END_IF;

    30:
        IF SensorWeight THEN
            AutoStep := 40;
        END_IF;

    40:
        IF weightEdge THEN
            tmp_unqualified := (weight < 100.0) OR (weight > 200.0);
            IF tmp_unqualified THEN
                kick := TRUE;
                AutoStep := 0;
            ELSE
                lastFiringTemp := 500.0 + (weight - 100.0) * 0.5;
                AutoStep := 50;
            END_IF;
        END_IF;

    50:
        IF SensorFiring THEN
            AutoStep := 60;
        END_IF;

    60:
        IF firingEdge THEN
            AutoStep := 70;
        END_IF;

    70:
        IF SensorOutput THEN
            AutoStep := 80;
        END_IF;

    80:
        IF NOT SensorOutput THEN
            AutoStep := 0;
        END_IF;
END_CASE;

MotorForward := (AutoStep = 10) OR (AutoStep = 30) OR (AutoStep = 50) OR (AutoStep = 70);
MotorReverse := FALSE;
CompletionLight := SensorOutput;
firingTemp := lastFiringTemp;
END_FUNCTION_BLOCK

(* ---- public-hard-06.raw_candidate_01.st ---- *)
FUNCTION_BLOCK ProductionControl
VAR_INPUT
    Mode : BOOL;
    ForwardButton : BOOL;
    ReverseButton : BOOL;
    SensorFeed : BOOL;
    SensorWash : BOOL;
    SensorWeight : BOOL;
    SensorFiring : BOOL;
    SensorOutput : BOOL;
    washComplete : BOOL;
    weightComplete : BOOL;
    weight : REAL;
    firingComplete : BOOL;
END_VAR
VAR_OUTPUT
    MotorForward : BOOL;
    MotorReverse : BOOL;
    kick : BOOL;
    CompletionLight : BOOL;
    firingTemp : REAL;
END_VAR
VAR
    AutoStep : INT := 0;
    AutoInit : BOOL := FALSE;
    lastFiringTemp : REAL := 0.0;
    rtWash : R_TRIG;
    rtWeight : R_TRIG;
    rtFiring : R_TRIG;
    washEdge : BOOL;
    weightEdge : BOOL;
    firingEdge : BOOL;
    tmp_unqualified : BOOL;
END_VAR

(*
ENGINEERING_CONTRACT
MotorForward: auto active in states 10/30/50/70; manual = ForwardButton AND NOT ReverseButton.
MotorReverse: manual only, interlocked with ForwardButton; both false if both buttons true.
kick: pulse on rising weightComplete when weight < 100 or weight > 200 (unqualified).
CompletionLight: combinational = SensorOutput while Mode=TRUE; off in manual.
firingTemp: stored on qualified weightComplete; formula 500 + (weight-100)*0.5, retained otherwise.
Units: weight REAL in same unit as thresholds; firingTemp REAL degrees; boundaries inclusive 100..200.
*)
(* CONTRACT_RULES [] *)

rtWash(CLK := washComplete);
rtWeight(CLK := weightComplete);
rtFiring(CLK := firingComplete);
washEdge := rtWash.Q;
weightEdge := rtWeight.Q;
firingEdge := rtFiring.Q;

IF NOT AutoInit THEN
    AutoInit := TRUE;
    IF SensorOutput THEN
        AutoStep := 80;
    ELSIF SensorFiring THEN
        AutoStep := 60;
    ELSIF SensorWeight THEN
        AutoStep := 40;
    ELSIF SensorWash THEN
        AutoStep := 20;
    ELSIF SensorFeed THEN
        AutoStep := 10;
    ELSE
        AutoStep := 0;
    END_IF;
END_IF;

IF NOT Mode THEN
    MotorForward := ForwardButton AND (NOT ReverseButton);
    MotorReverse := ReverseButton AND (NOT ForwardButton);
    kick := FALSE;
    CompletionLight := FALSE;
    firingTemp := lastFiringTemp;
    RETURN;
END_IF;

MotorForward := FALSE;
MotorReverse := FALSE;
kick := FALSE;
CompletionLight := FALSE;

CASE AutoStep OF
    0:
        IF SensorFeed THEN
            AutoStep := 10;
        END_IF;

    10:
        IF SensorWash THEN
            AutoStep := 20;
        END_IF;

    20:
        IF washEdge THEN
            AutoStep := 30;
        END_IF;

    30:
        IF SensorWeight THEN
            AutoStep := 40;
        END_IF;

    40:
        IF weightEdge THEN
            tmp_unqualified := (weight < 100.0) OR (weight > 200.0);
            IF tmp_unqualified THEN
                kick := TRUE;
                AutoStep := 0;
            ELSE
                lastFiringTemp := 500.0 + (weight - 100.0) * 0.5;
                AutoStep := 50;
            END_IF;
        END_IF;

    50:
        IF SensorFiring THEN
            AutoStep := 60;
        END_IF;

    60:
        IF firingEdge THEN
            AutoStep := 70;
        END_IF;

    70:
        IF SensorOutput THEN
            AutoStep := 80;
        END_IF;

    80:
        ;
END_CASE;

MotorForward := (AutoStep = 10) OR (AutoStep = 30) OR (AutoStep = 50) OR (AutoStep = 70);
MotorReverse := FALSE;
CompletionLight := SensorOutput;
firingTemp := lastFiringTemp;
END_FUNCTION_BLOCK

(* ---- public-hard-06.raw_candidate_02.st ---- *)
FUNCTION_BLOCK ProductionControl
VAR_INPUT
    Mode : BOOL;
    ForwardButton : BOOL;
    ReverseButton : BOOL;
    SensorFeed : BOOL;
    SensorWash : BOOL;
    SensorWeight : BOOL;
    SensorFiring : BOOL;
    SensorOutput : BOOL;
    washComplete : BOOL;
    weightComplete : BOOL;
    weight : REAL;
    firingComplete : BOOL;
END_VAR
VAR_OUTPUT
    MotorForward : BOOL;
    MotorReverse : BOOL;
    kick : BOOL;
    CompletionLight : BOOL;
    firingTemp : REAL;
END_VAR
VAR
    AutoStep : INT := 0;
    AutoInit : BOOL := FALSE;
    lastFiringTemp : REAL := 0.0;
    rtWash : R_TRIG;
    rtWeight : R_TRIG;
    rtFiring : R_TRIG;
    washEdge : BOOL;
    weightEdge : BOOL;
    firingEdge : BOOL;
    tmp_unqualified : BOOL;
END_VAR

(*
ENGINEERING_CONTRACT
MotorForward: auto active in states 10/30/50/70; manual = ForwardButton AND NOT ReverseButton.
MotorReverse: manual only, interlocked with ForwardButton; both false if both buttons true.
kick: pulse on rising weightComplete when weight < 100 or weight > 200 (unqualified).
CompletionLight: combinational = SensorOutput while Mode=TRUE; off in manual.
firingTemp: stored on qualified weightComplete; formula 500 + (weight-100)*0.5, retained otherwise.
Units: weight REAL in same unit as thresholds; firingTemp REAL degrees; boundaries inclusive 100..200.
*)
(* CONTRACT_RULES [] *)

rtWash(CLK := washComplete);
rtWeight(CLK := weightComplete);
rtFiring(CLK := firingComplete);
washEdge := rtWash.Q;
weightEdge := rtWeight.Q;
firingEdge := rtFiring.Q;

IF NOT AutoInit THEN
    AutoInit := TRUE;
    IF SensorOutput THEN
        AutoStep := 80;
    ELSIF SensorFiring THEN
        AutoStep := 60;
    ELSIF SensorWeight THEN
        AutoStep := 40;
    ELSIF SensorWash THEN
        AutoStep := 20;
    ELSIF SensorFeed THEN
        AutoStep := 10;
    ELSE
        AutoStep := 0;
    END_IF;
END_IF;

IF NOT Mode THEN
    MotorForward := ForwardButton AND (NOT ReverseButton);
    MotorReverse := ReverseButton AND (NOT ForwardButton);
    kick := FALSE;
    CompletionLight := FALSE;
    firingTemp := lastFiringTemp;
    RETURN;
END_IF;

MotorForward := FALSE;
MotorReverse := FALSE;
kick := FALSE;
CompletionLight := FALSE;

CASE AutoStep OF
    0:
        IF SensorFeed THEN
            AutoStep := 10;
        END_IF;

    10:
        IF SensorWash THEN
            AutoStep := 20;
        END_IF;

    20:
        IF washEdge THEN
            AutoStep := 30;
        END_IF;

    30:
        IF SensorWeight THEN
            AutoStep := 40;
        END_IF;

    40:
        IF weightEdge THEN
            tmp_unqualified := (weight < 100.0) OR (weight > 200.0);
            IF tmp_unqualified THEN
                kick := TRUE;
                AutoStep := 0;
            ELSE
                lastFiringTemp := 500.0 + (weight - 100.0) * 0.5;
                AutoStep := 50;
            END_IF;
        END_IF;

    50:
        IF SensorFiring THEN
            AutoStep := 60;
        END_IF;

    60:
        IF firingEdge THEN
            AutoStep := 70;
        END_IF;

    70:
        IF SensorOutput THEN
            AutoStep := 80;
        END_IF;

    80:
        IF NOT SensorOutput THEN
            AutoStep := 0;
        END_IF;
END_CASE;

MotorForward := (AutoStep = 10) OR (AutoStep = 30) OR (AutoStep = 50) OR (AutoStep = 70);
MotorReverse := FALSE;
CompletionLight := SensorOutput;
firingTemp := lastFiringTemp;
END_FUNCTION_BLOCK

(* ---- public-hard-06.raw_candidate_03.st ---- *)
FUNCTION_BLOCK ProductionControl
VAR_INPUT
    Mode : BOOL;
    ForwardButton : BOOL;
    ReverseButton : BOOL;
    SensorFeed : BOOL;
    SensorWash : BOOL;
    SensorWeight : BOOL;
    SensorFiring : BOOL;
    SensorOutput : BOOL;
    washComplete : BOOL;
    weightComplete : BOOL;
    weight : REAL;
    firingComplete : BOOL;
END_VAR
VAR_OUTPUT
    MotorForward : BOOL;
    MotorReverse : BOOL;
    kick : BOOL;
    CompletionLight : BOOL;
    firingTemp : REAL;
END_VAR
VAR
    AutoStep : INT := 0;
    AutoInit : BOOL := FALSE;
    lastFiringTemp : REAL := 0.0;
    rtWash : R_TRIG;
    rtWeight : R_TRIG;
    rtFiring : R_TRIG;
    washEdge : BOOL;
    weightEdge : BOOL;
    firingEdge : BOOL;
    rtMode : R_TRIG;
    ModeRise : BOOL;
    tmp_unqualified : BOOL;
END_VAR

(*
ENGINEERING_CONTRACT
MotorForward: auto active in states 10/30/50/70; manual = ForwardButton AND NOT ReverseButton.
MotorReverse: manual only, interlocked with ForwardButton; both false if both buttons true.
kick: pulse on rising weightComplete when weight < 100 or weight > 200 (unqualified).
CompletionLight: combinational = SensorOutput while Mode=TRUE; off in manual.
firingTemp: stored on qualified weightComplete; formula 500 + (weight-100)*0.5, retained otherwise.
Units: weight REAL in same unit as thresholds; firingTemp REAL degrees; boundaries inclusive 100..200.
*)
(* CONTRACT_RULES [] *)

rtMode(CLK := Mode);
ModeRise := rtMode.Q;
rtWash(CLK := washComplete);
rtWeight(CLK := weightComplete);
rtFiring(CLK := firingComplete);
washEdge := rtWash.Q;
weightEdge := rtWeight.Q;
firingEdge := rtFiring.Q;

IF (NOT AutoInit) OR ModeRise THEN
    AutoInit := TRUE;
    IF SensorOutput THEN
        AutoStep := 80;
    ELSIF SensorFiring THEN
        AutoStep := 60;
    ELSIF SensorWeight THEN
        AutoStep := 40;
    ELSIF SensorWash THEN
        AutoStep := 20;
    ELSIF SensorFeed THEN
        AutoStep := 10;
    ELSE
        AutoStep := 0;
    END_IF;
END_IF;

IF NOT Mode THEN
    MotorForward := ForwardButton AND (NOT ReverseButton);
    MotorReverse := ReverseButton AND (NOT ForwardButton);
    kick := FALSE;
    CompletionLight := FALSE;
    firingTemp := lastFiringTemp;
    RETURN;
END_IF;

MotorForward := FALSE;
MotorReverse := FALSE;
kick := FALSE;
CompletionLight := FALSE;

CASE AutoStep OF
    0:
        IF SensorFeed THEN
            AutoStep := 10;
        END_IF;

    10:
        IF SensorWash THEN
            AutoStep := 20;
        END_IF;

    20:
        IF washEdge THEN
            AutoStep := 30;
        END_IF;

    30:
        IF SensorWeight THEN
            AutoStep := 40;
        END_IF;

    40:
        IF weightEdge THEN
            tmp_unqualified := (weight < 100.0) OR (weight > 200.0);
            IF tmp_unqualified THEN
                kick := TRUE;
                AutoStep := 0;
            ELSE
                lastFiringTemp := 500.0 + (weight - 100.0) * 0.5;
                AutoStep := 50;
            END_IF;
        END_IF;

    50:
        IF SensorFiring THEN
            AutoStep := 60;
        END_IF;

    60:
        IF firingEdge THEN
            AutoStep := 70;
        END_IF;

    70:
        IF SensorOutput THEN
            AutoStep := 80;
        END_IF;

    80:
        IF NOT SensorOutput THEN
            AutoStep := 0;
        END_IF;
END_CASE;

MotorForward := (AutoStep = 10) OR (AutoStep = 30) OR (AutoStep = 50) OR (AutoStep = 70);
MotorReverse := FALSE;
CompletionLight := SensorOutput;
firingTemp := lastFiringTemp;
END_FUNCTION_BLOCK

(* ---- public-hard-06.raw_candidate_04.st ---- *)
FUNCTION_BLOCK ProductionControl
VAR_INPUT
    Mode : BOOL;
    ForwardButton : BOOL;
    ReverseButton : BOOL;
    SensorFeed : BOOL;
    SensorWash : BOOL;
    SensorWeight : BOOL;
    SensorFiring : BOOL;
    SensorOutput : BOOL;
    washComplete : BOOL;
    weightComplete : BOOL;
    weight : REAL;
    firingComplete : BOOL;
END_VAR
VAR_OUTPUT
    MotorForward : BOOL;
    MotorReverse : BOOL;
    kick : BOOL;
    CompletionLight : BOOL;
    firingTemp : REAL;
END_VAR
VAR
    AutoStep : INT := 0;
    AutoInit : BOOL := FALSE;
    lastFiringTemp : REAL := 0.0;
    rtWash : R_TRIG;
    rtWeight : R_TRIG;
    rtFiring : R_TRIG;
    washEdge : BOOL;
    weightEdge : BOOL;
    firingEdge : BOOL;
    rtMode : R_TRIG;
    ModeRise : BOOL;
    tmp_unqualified : BOOL;
END_VAR

(*
ENGINEERING_CONTRACT
MotorForward: auto active in states 10/30/50/70; manual = ForwardButton AND NOT ReverseButton.
MotorReverse: manual only, interlocked with ForwardButton; both false if both buttons true.
kick: pulse on rising weightComplete when weight < 100 or weight > 200 (unqualified).
CompletionLight: combinational = SensorOutput while Mode=TRUE; off in manual.
firingTemp: stored on qualified weightComplete; formula 500 + (weight-100)*0.5, retained otherwise.
Units: weight REAL in same unit as thresholds; firingTemp REAL degrees; boundaries inclusive 100..200.
*)
(* CONTRACT_RULES [] *)

rtMode(CLK := Mode);
ModeRise := rtMode.Q;
rtWash(CLK := washComplete);
rtWeight(CLK := weightComplete);
rtFiring(CLK := firingComplete);
washEdge := rtWash.Q;
weightEdge := rtWeight.Q;
firingEdge := rtFiring.Q;

IF (NOT AutoInit) OR ModeRise THEN
    AutoInit := TRUE;
    IF SensorOutput THEN
        AutoStep := 80;
    ELSIF SensorFiring THEN
        AutoStep := 60;
    ELSIF SensorWeight THEN
        AutoStep := 40;
    ELSIF SensorWash THEN
        AutoStep := 20;
    ELSIF SensorFeed THEN
        AutoStep := 10;
    ELSE
        AutoStep := 0;
    END_IF;
END_IF;

IF NOT Mode THEN
    MotorForward := ForwardButton AND (NOT ReverseButton);
    MotorReverse := ReverseButton AND (NOT ForwardButton);
    kick := FALSE;
    CompletionLight := FALSE;
    firingTemp := lastFiringTemp;
    RETURN;
END_IF;

MotorForward := FALSE;
MotorReverse := FALSE;
kick := FALSE;
CompletionLight := FALSE;

CASE AutoStep OF
    0:
        IF SensorFeed THEN
            AutoStep := 10;
        END_IF;

    10:
        IF SensorWash THEN
            AutoStep := 20;
        END_IF;

    20:
        IF washComplete THEN
            AutoStep := 30;
        END_IF;

    30:
        IF SensorWeight THEN
            AutoStep := 40;
        END_IF;

    40:
        IF weightComplete THEN
            tmp_unqualified := (weight < 100.0) OR (weight > 200.0);
            IF tmp_unqualified THEN
                kick := TRUE;
                AutoStep := 0;
            ELSE
                lastFiringTemp := 500.0 + (weight - 100.0) * 0.5;
                AutoStep := 50;
            END_IF;
        END_IF;

    50:
        IF SensorFiring THEN
            AutoStep := 60;
        END_IF;

    60:
        IF firingComplete THEN
            AutoStep := 70;
        END_IF;

    70:
        IF SensorOutput THEN
            AutoStep := 80;
        END_IF;

    80:
        IF NOT SensorOutput THEN
            AutoStep := 0;
        END_IF;
END_CASE;

MotorForward := (AutoStep = 10) OR (AutoStep = 30) OR (AutoStep = 50) OR (AutoStep = 70);
MotorReverse := FALSE;
CompletionLight := SensorOutput;
firingTemp := lastFiringTemp;
END_FUNCTION_BLOCK

(* ---- public-medium-01.candidate_01.st ---- *)
TYPE ST_Pump :
STRUCT
    priority : INT;
    selection : BOOL;
    RunComd : BOOL;
END_STRUCT
END_TYPE;

FUNCTION_BLOCK MultiPumpSwitchingControl
VAR_INPUT
    mode : BOOL;
    start : BOOL;
    stop : BOOL;
END_VAR
VAR_IN_OUT
    pumpGroup : ARRAY[1..5] OF ST_Pump;
END_VAR
VAR
    running : BOOL := FALSE;
    tmp_startPrev : BOOL := FALSE;
    tmp_i : INT;
    tmp_j : INT;
    tmp_k : INT;
    tmp_order : ARRAY[1..5] OF INT;
    tmp_isTop : ARRAY[1..5] OF BOOL;
    tmp_prioLeft : INT;
    tmp_prioRight : INT;
END_VAR

(* ENGINEERING_CONTRACT
- Mode select: PUB001/PUB003. mode FALSE=manual, TRUE=auto; outputs follow current mode each scan.
- Running latch: rising edge of start (PUB002) sets running=TRUE; stop=TRUE (PUB004) resets running=FALSE.
- Same-scan priority: stop overrides start; stop and start tests use final same-scan input values.
- Manual RunComd (PUB001/PUB003): RunComd[i] = running AND pumpGroup[i].selection, i=1..5.
- Auto RunComd (PUB001/PUB002): top 3 priorities selected each scan; larger priority wins.
  Ties are unspecified; this block breaks ties by lower array index.
  RunComd[i] = running AND tmp_isTop[i].
- Running state is retained across mode changes until stop; no unstated mode-change reset.
- Units/boundaries: array indices 1..5, priority INT, RunComd BOOL.
*)
(* CONTRACT_RULES [] *)

IF stop THEN
    running := FALSE;
ELSIF (NOT tmp_startPrev) AND start THEN
    running := TRUE;
END_IF;

tmp_startPrev := start;

IF NOT mode THEN
    FOR tmp_i := 1 TO 5 DO
        pumpGroup[tmp_i].RunComd := running AND pumpGroup[tmp_i].selection;
    END_FOR;
ELSE
    FOR tmp_i := 1 TO 5 DO
        tmp_order[tmp_i] := tmp_i;
        tmp_isTop[tmp_i] := FALSE;
    END_FOR;

    FOR tmp_i := 1 TO 4 DO
        FOR tmp_j := tmp_i + 1 TO 5 DO
            tmp_prioRight := pumpGroup[tmp_order[tmp_j]].priority;
            tmp_prioLeft := pumpGroup[tmp_order[tmp_i]].priority;
            IF tmp_prioRight > tmp_prioLeft THEN
                tmp_k := tmp_order[tmp_i];
                tmp_order[tmp_i] := tmp_order[tmp_j];
                tmp_order[tmp_j] := tmp_k;
            END_IF;
        END_FOR;
    END_FOR;

    FOR tmp_i := 1 TO 3 DO
        tmp_isTop[tmp_order[tmp_i]] := TRUE;
    END_FOR;

    FOR tmp_i := 1 TO 5 DO
        pumpGroup[tmp_i].RunComd := running AND tmp_isTop[tmp_i];
    END_FOR;
END_IF;

END_FUNCTION_BLOCK

(* ---- public-medium-01.candidate_02.st ---- *)
TYPE ST_Pump :
STRUCT
    priority : INT;
    selection : BOOL;
    RunComd : BOOL;
END_STRUCT
END_TYPE;

FUNCTION_BLOCK MultiPumpSwitchingControl
VAR_INPUT
    mode : BOOL;
    start : BOOL;
    stop : BOOL;
END_VAR
VAR_IN_OUT
    pumpGroup : ARRAY[1..5] OF ST_Pump;
END_VAR
VAR
    running : BOOL := FALSE;
    tmp_i : INT;
    tmp_j : INT;
    tmp_k : INT;
    tmp_order : ARRAY[1..5] OF INT;
    tmp_isTop : ARRAY[1..5] OF BOOL;
    tmp_prioLeft : INT;
    tmp_prioRight : INT;
END_VAR

(* ENGINEERING_CONTRACT
- Mode select: PUB001/PUB003. mode FALSE=manual, TRUE=auto; outputs follow current mode each scan.
- Running latch: level-sensitive set/reset. stop=TRUE (PUB004) resets running=FALSE; otherwise start=TRUE (PUB002) sets running=TRUE. Once set, running remains TRUE until stop even if start goes FALSE.
- Same-scan priority: stop overrides start; stop and start tests use final same-scan input values.
- Manual RunComd (PUB001/PUB003): RunComd[i] = running AND pumpGroup[i].selection, i=1..5.
- Auto RunComd (PUB001/PUB002): top 3 priorities selected each scan; larger priority wins.
  Ties are unspecified; this block breaks ties by lower array index.
  RunComd[i] = running AND tmp_isTop[i].
- Running state is retained across mode changes until stop; no unstated mode-change reset.
- Units/boundaries: array indices 1..5, priority INT, RunComd BOOL.
*)
(* CONTRACT_RULES [] *)

IF stop THEN
    running := FALSE;
ELSIF start THEN
    running := TRUE;
END_IF;

IF NOT mode THEN
    FOR tmp_i := 1 TO 5 DO
        pumpGroup[tmp_i].RunComd := running AND pumpGroup[tmp_i].selection;
    END_FOR;
ELSE
    FOR tmp_i := 1 TO 5 DO
        tmp_order[tmp_i] := tmp_i;
        tmp_isTop[tmp_i] := FALSE;
    END_FOR;

    FOR tmp_i := 1 TO 4 DO
        FOR tmp_j := tmp_i + 1 TO 5 DO
            tmp_prioRight := pumpGroup[tmp_order[tmp_j]].priority;
            tmp_prioLeft := pumpGroup[tmp_order[tmp_i]].priority;
            IF tmp_prioRight > tmp_prioLeft THEN
                tmp_k := tmp_order[tmp_i];
                tmp_order[tmp_i] := tmp_order[tmp_j];
                tmp_order[tmp_j] := tmp_k;
            END_IF;
        END_FOR;
    END_FOR;

    FOR tmp_i := 1 TO 3 DO
        tmp_isTop[tmp_order[tmp_i]] := TRUE;
    END_FOR;

    FOR tmp_i := 1 TO 5 DO
        pumpGroup[tmp_i].RunComd := running AND tmp_isTop[tmp_i];
    END_FOR;
END_IF;

END_FUNCTION_BLOCK

(* ---- public-medium-01.patch_base_02.st ---- *)
TYPE ST_Pump :
STRUCT
    priority : INT;
    selection : BOOL;
    RunComd : BOOL;
END_STRUCT
END_TYPE;

FUNCTION_BLOCK MultiPumpSwitchingControl
VAR_INPUT
    mode : BOOL;
    start : BOOL;
    stop : BOOL;
END_VAR
VAR_IN_OUT
    pumpGroup : ARRAY[1..5] OF ST_Pump;
END_VAR
VAR
    running : BOOL := FALSE;
    tmp_startPrev : BOOL := FALSE;
    tmp_i : INT;
    tmp_j : INT;
    tmp_k : INT;
    tmp_order : ARRAY[1..5] OF INT;
    tmp_isTop : ARRAY[1..5] OF BOOL;
    tmp_prioLeft : INT;
    tmp_prioRight : INT;
END_VAR

(* ENGINEERING_CONTRACT
- Mode select: PUB001/PUB003. mode FALSE=manual, TRUE=auto; outputs follow current mode each scan.
- Running latch: rising edge of start (PUB002) sets running=TRUE; stop=TRUE (PUB004) resets running=FALSE.
- Same-scan priority: stop overrides start; stop and start tests use final same-scan input values.
- Manual RunComd (PUB001/PUB003): RunComd[i] = running AND pumpGroup[i].selection, i=1..5.
- Auto RunComd (PUB001/PUB002): top 3 priorities selected each scan; larger priority wins.
  Ties are unspecified; this block breaks ties by lower array index.
  RunComd[i] = running AND tmp_isTop[i].
- Running state is retained across mode changes until stop; no unstated mode-change reset.
- Units/boundaries: array indices 1..5, priority INT, RunComd BOOL.
*)
(* CONTRACT_RULES [] *)

IF stop THEN
    running := FALSE;
ELSIF (NOT tmp_startPrev) AND start THEN
    running := TRUE;
END_IF;

tmp_startPrev := start;

IF NOT mode THEN
    FOR tmp_i := 1 TO 5 DO
        pumpGroup[tmp_i].RunComd := running AND pumpGroup[tmp_i].selection;
    END_FOR;
ELSE
    FOR tmp_i := 1 TO 5 DO
        tmp_order[tmp_i] := tmp_i;
        tmp_isTop[tmp_i] := FALSE;
    END_FOR;

    FOR tmp_i := 1 TO 4 DO
        FOR tmp_j := tmp_i + 1 TO 5 DO
            tmp_prioRight := pumpGroup[tmp_order[tmp_j]].priority;
            tmp_prioLeft := pumpGroup[tmp_order[tmp_i]].priority;
            IF tmp_prioRight > tmp_prioLeft THEN
                tmp_k := tmp_order[tmp_i];
                tmp_order[tmp_i] := tmp_order[tmp_j];
                tmp_order[tmp_j] := tmp_k;
            END_IF;
        END_FOR;
    END_FOR;

    FOR tmp_i := 1 TO 3 DO
        tmp_isTop[tmp_order[tmp_i]] := TRUE;
    END_FOR;

    FOR tmp_i := 1 TO 5 DO
        pumpGroup[tmp_i].RunComd := running AND tmp_isTop[tmp_i];
    END_FOR;
END_IF;

END_FUNCTION_BLOCK

(* ---- public-medium-01.raw_candidate_01.st ---- *)
TYPE ST_Pump :
STRUCT
    priority : INT;
    selection : BOOL;
    RunComd : BOOL;
END_STRUCT
END_TYPE

FUNCTION_BLOCK MultiPumpSwitchingControl
VAR_INPUT
    mode : BOOL;
    start : BOOL;
    stop : BOOL;
END_VAR
VAR_IN_OUT
    pumpGroup : ARRAY[1..5] OF ST_Pump;
END_VAR
VAR
    running : BOOL := FALSE;
    tmp_startPrev : BOOL := FALSE;
    tmp_i : INT;
    tmp_j : INT;
    tmp_k : INT;
    tmp_order : ARRAY[1..5] OF INT;
    tmp_isTop : ARRAY[1..5] OF BOOL;
    tmp_prioLeft : INT;
    tmp_prioRight : INT;
END_VAR

(* ENGINEERING_CONTRACT
- Mode select: PUB001/PUB003. mode FALSE=manual, TRUE=auto; outputs follow current mode each scan.
- Running latch: rising edge of start (PUB002) sets running=TRUE; stop=TRUE (PUB004) resets running=FALSE.
- Same-scan priority: stop overrides start; stop and start tests use final same-scan input values.
- Manual RunComd (PUB001/PUB003): RunComd[i] = running AND pumpGroup[i].selection, i=1..5.
- Auto RunComd (PUB001/PUB002): top 3 priorities selected each scan; larger priority wins.
  Ties are unspecified; this block breaks ties by lower array index.
  RunComd[i] = running AND tmp_isTop[i].
- Running state is retained across mode changes until stop; no unstated mode-change reset.
- Units/boundaries: array indices 1..5, priority INT, RunComd BOOL.
*)
(* CONTRACT_RULES [] *)

IF stop THEN
    running := FALSE;
ELSIF (NOT tmp_startPrev) AND start THEN
    running := TRUE;
END_IF;

tmp_startPrev := start;

IF NOT mode THEN
    FOR tmp_i := 1 TO 5 DO
        pumpGroup[tmp_i].RunComd := running AND pumpGroup[tmp_i].selection;
    END_FOR;
ELSE
    FOR tmp_i := 1 TO 5 DO
        tmp_order[tmp_i] := tmp_i;
        tmp_isTop[tmp_i] := FALSE;
    END_FOR;

    FOR tmp_i := 1 TO 4 DO
        FOR tmp_j := tmp_i + 1 TO 5 DO
            tmp_prioRight := pumpGroup[tmp_order[tmp_j]].priority;
            tmp_prioLeft := pumpGroup[tmp_order[tmp_i]].priority;
            IF tmp_prioRight > tmp_prioLeft THEN
                tmp_k := tmp_order[tmp_i];
                tmp_order[tmp_i] := tmp_order[tmp_j];
                tmp_order[tmp_j] := tmp_k;
            END_IF;
        END_FOR;
    END_FOR;

    FOR tmp_i := 1 TO 3 DO
        tmp_isTop[tmp_order[tmp_i]] := TRUE;
    END_FOR;

    FOR tmp_i := 1 TO 5 DO
        pumpGroup[tmp_i].RunComd := running AND tmp_isTop[tmp_i];
    END_FOR;
END_IF;

END_FUNCTION_BLOCK

(* ---- public-medium-01.raw_candidate_02.st ---- *)
TYPE ST_Pump :
STRUCT
    priority : INT;
    selection : BOOL;
    RunComd : BOOL;
END_STRUCT
END_TYPE;

FUNCTION_BLOCK MultiPumpSwitchingControl
VAR_INPUT
    mode : BOOL;
    start : BOOL;
    stop : BOOL;
END_VAR
VAR_IN_OUT
    pumpGroup : ARRAY[1..5] OF ST_Pump;
END_VAR
VAR
    running : BOOL := FALSE;
    tmp_i : INT;
    tmp_j : INT;
    tmp_k : INT;
    tmp_order : ARRAY[1..5] OF INT;
    tmp_isTop : ARRAY[1..5] OF BOOL;
    tmp_prioLeft : INT;
    tmp_prioRight : INT;
END_VAR

(* ENGINEERING_CONTRACT
- Mode select: PUB001/PUB003. mode FALSE=manual, TRUE=auto; outputs follow current mode each scan.
- Running latch: level-sensitive set/reset. stop=TRUE (PUB004) resets running=FALSE; otherwise start=TRUE (PUB002) sets running=TRUE. Once set, running remains TRUE until stop even if start goes FALSE.
- Same-scan priority: stop overrides start; stop and start tests use final same-scan input values.
- Manual RunComd (PUB001/PUB003): RunComd[i] = running AND pumpGroup[i].selection, i=1..5.
- Auto RunComd (PUB001/PUB002): top 3 priorities selected each scan; larger priority wins.
  Ties are unspecified; this block breaks ties by lower array index.
  RunComd[i] = running AND tmp_isTop[i].
- Running state is retained across mode changes until stop; no unstated mode-change reset.
- Units/boundaries: array indices 1..5, priority INT, RunComd BOOL.
*)
(* CONTRACT_RULES [] *)

IF stop THEN
    running := FALSE;
ELSIF start THEN
    running := TRUE;
END_IF;

IF NOT mode THEN
    FOR tmp_i := 1 TO 5 DO
        pumpGroup[tmp_i].RunComd := running AND pumpGroup[tmp_i].selection;
    END_FOR;
ELSE
    FOR tmp_i := 1 TO 5 DO
        tmp_order[tmp_i] := tmp_i;
        tmp_isTop[tmp_i] := FALSE;
    END_FOR;

    FOR tmp_i := 1 TO 4 DO
        FOR tmp_j := tmp_i + 1 TO 5 DO
            tmp_prioRight := pumpGroup[tmp_order[tmp_j]].priority;
            tmp_prioLeft := pumpGroup[tmp_order[tmp_i]].priority;
            IF tmp_prioRight > tmp_prioLeft THEN
                tmp_k := tmp_order[tmp_i];
                tmp_order[tmp_i] := tmp_order[tmp_j];
                tmp_order[tmp_j] := tmp_k;
            END_IF;
        END_FOR;
    END_FOR;

    FOR tmp_i := 1 TO 3 DO
        tmp_isTop[tmp_order[tmp_i]] := TRUE;
    END_FOR;

    FOR tmp_i := 1 TO 5 DO
        pumpGroup[tmp_i].RunComd := running AND tmp_isTop[tmp_i];
    END_FOR;
END_IF;

END_FUNCTION_BLOCK

(* ---- public-medium-02.candidate_01.st ---- *)
TYPE ST_AnalogChannel :
STRUCT
    enable : BOOL;
    hiLIM : REAL;
    loLIM : REAL;
    bipolar : BOOL;
    measuringMode : INT;
    retVal : WORD;
    outputValue : REAL;
END_STRUCT
END_TYPE;

(* ENGINEERING_CONTRACT
   Loop count: count limited to 0..min(array lengths); ordinal start at each array lower bound (PUB001).
   channels[].retVal: activated on enabled scan; invalid mode -> 16#8001, invalid limits -> 16#8002,
   success -> 0 (PUB006, PUB007, PUB008).
   channels[].outputValue: written only on successful conversion; mode 0 linear scaling,
   mode 1 /10, mode 2 /100 (PUB003, PUB004, PUB005).
   Disabled channels retain prior retVal/outputValue (unspecified retention interpretation).
*)

(* CONTRACT_RULES [] *)

FUNCTION_BLOCK AnalogBatchProcessing
VAR_INPUT
    count : DINT;
END_VAR
VAR_IN_OUT
    analogValues : ARRAY[*] OF INT;
    channels : ARRAY[*] OF ST_AnalogChannel;
END_VAR
VAR
    local_i : DINT;
    local_n : DINT;
    local_analog_idx : DINT;
    local_channel_idx : DINT;
    local_raw : INT;
    local_mode : INT;
    local_min_len : DINT;
    local_ch_len : DINT;
    local_raw_min : REAL;
    local_raw_max : REAL;
    local_span_raw : REAL;
    local_ratio : REAL;
END_VAR

local_n := count;
IF local_n < 0 THEN
    local_n := 0;
END_IF;

local_min_len := UPPER_BOUND(analogValues, 1) - LOWER_BOUND(analogValues, 1) + 1;
local_ch_len := UPPER_BOUND(channels, 1) - LOWER_BOUND(channels, 1) + 1;
IF local_min_len > local_ch_len THEN
    local_min_len := local_ch_len;
END_IF;
IF local_n > local_min_len THEN
    local_n := local_min_len;
END_IF;

IF local_n > 0 THEN
    FOR local_i := 0 TO local_n - 1 DO
        local_analog_idx := LOWER_BOUND(analogValues, 1) + local_i;
        local_channel_idx := LOWER_BOUND(channels, 1) + local_i;

        IF channels[local_channel_idx].enable THEN
            local_mode := channels[local_channel_idx].measuringMode;

            IF (local_mode <> 0) AND (local_mode <> 1) AND (local_mode <> 2) THEN
                channels[local_channel_idx].retVal := 16#8001;
                (* skip conversion: outputValue unchanged *)
            ELSIF channels[local_channel_idx].hiLIM <= channels[local_channel_idx].loLIM THEN
                channels[local_channel_idx].retVal := 16#8002;
                (* skip conversion: outputValue unchanged *)
            ELSE
                channels[local_channel_idx].retVal := 0;
                CASE local_mode OF
                    0:
                        local_raw := analogValues[local_analog_idx];
                        IF channels[local_channel_idx].bipolar THEN
                            local_raw_min := -27648.0;
                            local_raw_max := 27648.0;
                        ELSE
                            local_raw_min := 0.0;
                            local_raw_max := 27648.0;
                        END_IF;

                        local_span_raw := local_raw_max - local_raw_min;
                        local_ratio := (TO_REAL(local_raw) - local_raw_min) / local_span_raw;
                        channels[local_channel_idx].outputValue := channels[local_channel_idx].loLIM
                            + local_ratio * (channels[local_channel_idx].hiLIM - channels[local_channel_idx].loLIM);

                    1:
                        channels[local_channel_idx].outputValue := TO_REAL(analogValues[local_analog_idx]) / 10.0;

                    2:
                        channels[local_channel_idx].outputValue := TO_REAL(analogValues[local_analog_idx]) / 100.0;
                END_CASE;
            END_IF;
        ELSE
            (* disabled: no writes to retVal or outputValue *)
        END_IF;
    END_FOR;
END_IF;

(* ---- public-medium-02.candidate_02.st ---- *)
TYPE ST_AnalogChannel :
STRUCT
    enable : BOOL;
    hiLIM : REAL;
    loLIM : REAL;
    bipolar : BOOL;
    measuringMode : INT;
    retVal : WORD;
    outputValue : REAL;
END_STRUCT
END_TYPE;

(* ENGINEERING_CONTRACT
   Loop count: count limited to 0..min(array lengths); ordinal start at each array lower bound (PUB001).
   channels[].retVal: activated on enabled scan; invalid mode -> 16#8001, invalid limits -> 16#8002,
   success -> 0 (PUB006, PUB007, PUB008).
   channels[].outputValue: written only on successful conversion; mode 0 linear scaling,
   mode 1 /10, mode 2 /100 (PUB003, PUB004, PUB005).
   Disabled channels retain prior retVal/outputValue (unspecified retention interpretation).
*)

(* CONTRACT_RULES [] *)

FUNCTION_BLOCK AnalogBatchProcessing
VAR_INPUT
    count : DINT;
END_VAR
VAR_IN_OUT
    analogValues : ARRAY[*] OF INT;
    channels : ARRAY[*] OF ST_AnalogChannel;
END_VAR
VAR
    local_i : DINT;
    local_n : DINT;
    local_analog_idx : DINT;
    local_channel_idx : DINT;
    local_raw : INT;
    local_mode : INT;
    local_min_len : DINT;
    local_ch_len : DINT;
    local_raw_min : REAL;
    local_raw_max : REAL;
    local_span_raw : REAL;
    local_ratio : REAL;
END_VAR

local_n := count;
IF local_n < 0 THEN
    local_n := 0;
END_IF;

local_min_len := UPPER_BOUND(analogValues, 1) - LOWER_BOUND(analogValues, 1) + 1;
local_ch_len := UPPER_BOUND(channels, 1) - LOWER_BOUND(channels, 1) + 1;
IF local_min_len > local_ch_len THEN
    local_min_len := local_ch_len;
END_IF;
IF local_n > local_min_len THEN
    local_n := local_min_len;
END_IF;

IF local_n > 0 THEN
    FOR local_i := 0 TO local_n - 1 DO
        local_analog_idx := LOWER_BOUND(analogValues, 1) + local_i;
        local_channel_idx := LOWER_BOUND(channels, 1) + local_i;

        IF channels[local_channel_idx].enable THEN
            local_mode := channels[local_channel_idx].measuringMode;

            IF (local_mode <> 0) AND (local_mode <> 1) AND (local_mode <> 2) THEN
                channels[local_channel_idx].retVal := 16#8001;
                (* skip conversion: outputValue unchanged *)
            ELSIF channels[local_channel_idx].hiLIM <= channels[local_channel_idx].loLIM THEN
                channels[local_channel_idx].retVal := 16#8002;
                (* skip conversion: outputValue unchanged *)
            ELSE
                channels[local_channel_idx].retVal := 0;
                CASE local_mode OF
                    0:
                        local_raw := analogValues[local_analog_idx];
                        IF channels[local_channel_idx].bipolar THEN
                            local_raw_min := -27648.0;
                            local_raw_max := 27648.0;
                        ELSE
                            local_raw_min := 0.0;
                            local_raw_max := 27648.0;
                        END_IF;

                        local_span_raw := local_raw_max - local_raw_min;
                        local_ratio := (TO_REAL(local_raw) - local_raw_min) / local_span_raw;
                        channels[local_channel_idx].outputValue := channels[local_channel_idx].loLIM
                            + local_ratio * (channels[local_channel_idx].hiLIM - channels[local_channel_idx].loLIM);

                    1:
                        channels[local_channel_idx].outputValue := TO_REAL(analogValues[local_analog_idx]) / 10.0;

                    2:
                        channels[local_channel_idx].outputValue := TO_REAL(analogValues[local_analog_idx]) / 100.0;
                END_CASE;
            END_IF;
        ELSE
            (* disabled: no writes to retVal or outputValue *)
        END_IF;
    END_FOR;
END_IF;

END_FUNCTION_BLOCK

(* ---- public-medium-02.candidate_03.st ---- *)
TYPE ST_AnalogChannel :
STRUCT
    enable : BOOL;
    hiLIM : REAL;
    loLIM : REAL;
    bipolar : BOOL;
    measuringMode : INT;
    retVal : WORD;
    outputValue : REAL;
END_STRUCT
END_TYPE;

(* ENGINEERING_CONTRACT
   Loop count: count limited to 0..min(array lengths); ordinal start at each array lower bound (PUB001).
   channels[].retVal: activated on enabled scan; invalid mode -> 16#8001, invalid limits -> 16#8002,
   success -> 0 (PUB006, PUB007, PUB008).
   channels[].outputValue: written only on successful conversion; mode 0 linear scaling,
   mode 1 /10, mode 2 /100 (PUB003, PUB004, PUB005).
   Disabled channels retain prior retVal/outputValue (unspecified retention interpretation).
*)

(* CONTRACT_RULES [] *)

FUNCTION_BLOCK AnalogBatchProcessing
VAR_INPUT
    count : DINT;
END_VAR
VAR_IN_OUT
    analogValues : ARRAY[*] OF INT;
    channels : ARRAY[*] OF ST_AnalogChannel;
END_VAR
VAR
    local_i : DINT;
    local_n : DINT;
    local_analog_idx : DINT;
    local_channel_idx : DINT;
    local_raw : INT;
    local_mode : INT;
    local_min_len : DINT;
    local_ch_len : DINT;
    local_raw_min : REAL;
    local_raw_max : REAL;
    local_span_raw : REAL;
    local_ratio : REAL;
END_VAR

local_n := count;
IF local_n < 0 THEN
    local_n := 0;
END_IF;

local_min_len := UPPER_BOUND(analogValues, 1) - LOWER_BOUND(analogValues, 1) + 1;
local_ch_len := UPPER_BOUND(channels, 1) - LOWER_BOUND(channels, 1) + 1;
IF local_min_len > local_ch_len THEN
    local_min_len := local_ch_len;
END_IF;
IF local_n > local_min_len THEN
    local_n := local_min_len;
END_IF;

IF local_n > 0 THEN
    FOR local_i := 0 TO local_n - 1 DO
        local_analog_idx := LOWER_BOUND(analogValues, 1) + local_i;
        local_channel_idx := LOWER_BOUND(channels, 1) + local_i;

        IF channels[local_channel_idx].enable THEN
            local_mode := channels[local_channel_idx].measuringMode;

            IF (local_mode <> 0) AND (local_mode <> 1) AND (local_mode <> 2) THEN
                channels[local_channel_idx].retVal := 16#8001;
                (* skip conversion: outputValue unchanged *)
            ELSIF channels[local_channel_idx].hiLIM <= channels[local_channel_idx].loLIM THEN
                channels[local_channel_idx].retVal := 16#8002;
                (* skip conversion: outputValue unchanged *)
            ELSE
                channels[local_channel_idx].retVal := 0;
                CASE local_mode OF
                    0:
                        local_raw := analogValues[local_analog_idx];
                        IF channels[local_channel_idx].bipolar THEN
                            local_raw_min := -27648.0;
                            local_raw_max := 27648.0;
                        ELSE
                            local_raw_min := 0.0;
                            local_raw_max := 27648.0;
                        END_IF;

                        local_span_raw := local_raw_max - local_raw_min;
                        local_ratio := (TO_REAL(local_raw) - local_raw_min) / local_span_raw;
                        channels[local_channel_idx].outputValue := channels[local_channel_idx].loLIM
                            + local_ratio * (channels[local_channel_idx].hiLIM - channels[local_channel_idx].loLIM);

                    1:
                        channels[local_channel_idx].outputValue := TO_REAL(analogValues[local_analog_idx]) / 10.0;

                    2:
                        channels[local_channel_idx].outputValue := TO_REAL(analogValues[local_analog_idx]) / 100.0;
                END_CASE;
            END_IF;
        ELSE
            (* disabled: no writes to retVal or outputValue *)
        END_IF;
    END_FOR;
END_IF;

END_FUNCTION_BLOCK

(* ---- public-medium-02.patch_base_02.st ---- *)
TYPE ST_AnalogChannel :
STRUCT
    enable : BOOL;
    hiLIM : REAL;
    loLIM : REAL;
    bipolar : BOOL;
    measuringMode : INT;
    retVal : WORD;
    outputValue : REAL;
END_STRUCT
END_TYPE;

(* ENGINEERING_CONTRACT
   Loop count: count limited to 0..min(array lengths); ordinal start at each array lower bound (PUB001).
   channels[].retVal: activated on enabled scan; invalid mode -> 16#8001, invalid limits -> 16#8002,
   success -> 0 (PUB006, PUB007, PUB008).
   channels[].outputValue: written only on successful conversion; mode 0 linear scaling,
   mode 1 /10, mode 2 /100 (PUB003, PUB004, PUB005).
   Disabled channels retain prior retVal/outputValue (unspecified retention interpretation).
*)

(* CONTRACT_RULES [] *)

FUNCTION_BLOCK AnalogBatchProcessing
VAR_INPUT
    count : DINT;
END_VAR
VAR_IN_OUT
    analogValues : ARRAY[*] OF INT;
    channels : ARRAY[*] OF ST_AnalogChannel;
END_VAR
VAR
    local_i : DINT;
    local_n : DINT;
    local_analog_idx : DINT;
    local_channel_idx : DINT;
    local_raw : INT;
    local_mode : INT;
    local_min_len : DINT;
    local_ch_len : DINT;
    local_raw_min : REAL;
    local_raw_max : REAL;
    local_span_raw : REAL;
    local_ratio : REAL;
END_VAR

local_n := count;
IF local_n < 0 THEN
    local_n := 0;
END_IF;

local_min_len := UPPER_BOUND(analogValues, 1) - LOWER_BOUND(analogValues, 1) + 1;
local_ch_len := UPPER_BOUND(channels, 1) - LOWER_BOUND(channels, 1) + 1;
IF local_min_len > local_ch_len THEN
    local_min_len := local_ch_len;
END_IF;
IF local_n > local_min_len THEN
    local_n := local_min_len;
END_IF;

IF local_n > 0 THEN
    FOR local_i := 0 TO local_n - 1 DO
        local_analog_idx := LOWER_BOUND(analogValues, 1) + local_i;
        local_channel_idx := LOWER_BOUND(channels, 1) + local_i;

        IF channels[local_channel_idx].enable THEN
            local_mode := channels[local_channel_idx].measuringMode;

            IF (local_mode <> 0) AND (local_mode <> 1) AND (local_mode <> 2) THEN
                channels[local_channel_idx].retVal := 16#8001;
                (* skip conversion: outputValue unchanged *)
            ELSIF channels[local_channel_idx].hiLIM <= channels[local_channel_idx].loLIM THEN
                channels[local_channel_idx].retVal := 16#8002;
                (* skip conversion: outputValue unchanged *)
            ELSE
                channels[local_channel_idx].retVal := 0;
                CASE local_mode OF
                    0:
                        local_raw := analogValues[local_analog_idx];
                        IF channels[local_channel_idx].bipolar THEN
                            local_raw_min := -27648.0;
                            local_raw_max := 27648.0;
                        ELSE
                            local_raw_min := 0.0;
                            local_raw_max := 27648.0;
                        END_IF;

                        local_span_raw := local_raw_max - local_raw_min;
                        local_ratio := (TO_REAL(local_raw) - local_raw_min) / local_span_raw;
                        channels[local_channel_idx].outputValue := channels[local_channel_idx].loLIM
                            + local_ratio * (channels[local_channel_idx].hiLIM - channels[local_channel_idx].loLIM);

                    1:
                        channels[local_channel_idx].outputValue := TO_REAL(analogValues[local_analog_idx]) / 10.0;

                    2:
                        channels[local_channel_idx].outputValue := TO_REAL(analogValues[local_analog_idx]) / 100.0;
                END_CASE;
            END_IF;
        ELSE
            (* disabled: no writes to retVal or outputValue *)
        END_IF;
    END_FOR;
END_IF;

(* ---- public-medium-02.patch_base_03.st ---- *)
TYPE ST_AnalogChannel :
STRUCT
    enable : BOOL;
    hiLIM : REAL;
    loLIM : REAL;
    bipolar : BOOL;
    measuringMode : INT;
    retVal : WORD;
    outputValue : REAL;
END_STRUCT
END_TYPE;

(* ENGINEERING_CONTRACT
   Loop count: count limited to 0..min(array lengths); ordinal start at each array lower bound (PUB001).
   channels[].retVal: activated on enabled scan; invalid mode -> 16#8001, invalid limits -> 16#8002,
   success -> 0 (PUB006, PUB007, PUB008).
   channels[].outputValue: written only on successful conversion; mode 0 linear scaling,
   mode 1 /10, mode 2 /100 (PUB003, PUB004, PUB005).
   Disabled channels retain prior retVal/outputValue (unspecified retention interpretation).
*)

(* CONTRACT_RULES [] *)

FUNCTION_BLOCK AnalogBatchProcessing
VAR_INPUT
    count : DINT;
END_VAR
VAR_IN_OUT
    analogValues : ARRAY[*] OF INT;
    channels : ARRAY[*] OF ST_AnalogChannel;
END_VAR
VAR
    local_i : DINT;
    local_n : DINT;
    local_analog_idx : DINT;
    local_channel_idx : DINT;
    local_raw : INT;
    local_mode : INT;
    local_min_len : DINT;
    local_ch_len : DINT;
    local_raw_min : REAL;
    local_raw_max : REAL;
    local_span_raw : REAL;
    local_ratio : REAL;
END_VAR

local_n := count;
IF local_n < 0 THEN
    local_n := 0;
END_IF;

local_min_len := UPPER_BOUND(analogValues, 1) - LOWER_BOUND(analogValues, 1) + 1;
local_ch_len := UPPER_BOUND(channels, 1) - LOWER_BOUND(channels, 1) + 1;
IF local_min_len > local_ch_len THEN
    local_min_len := local_ch_len;
END_IF;
IF local_n > local_min_len THEN
    local_n := local_min_len;
END_IF;

IF local_n > 0 THEN
    FOR local_i := 0 TO local_n - 1 DO
        local_analog_idx := LOWER_BOUND(analogValues, 1) + local_i;
        local_channel_idx := LOWER_BOUND(channels, 1) + local_i;

        IF channels[local_channel_idx].enable THEN
            local_mode := channels[local_channel_idx].measuringMode;

            IF (local_mode <> 0) AND (local_mode <> 1) AND (local_mode <> 2) THEN
                channels[local_channel_idx].retVal := 16#8001;
                (* skip conversion: outputValue unchanged *)
            ELSIF channels[local_channel_idx].hiLIM <= channels[local_channel_idx].loLIM THEN
                channels[local_channel_idx].retVal := 16#8002;
                (* skip conversion: outputValue unchanged *)
            ELSE
                channels[local_channel_idx].retVal := 0;
                CASE local_mode OF
                    0:
                        local_raw := analogValues[local_analog_idx];
                        IF channels[local_channel_idx].bipolar THEN
                            local_raw_min := -27648.0;
                            local_raw_max := 27648.0;
                        ELSE
                            local_raw_min := 0.0;
                            local_raw_max := 27648.0;
                        END_IF;

                        local_span_raw := local_raw_max - local_raw_min;
                        local_ratio := (TO_REAL(local_raw) - local_raw_min) / local_span_raw;
                        channels[local_channel_idx].outputValue := channels[local_channel_idx].loLIM
                            + local_ratio * (channels[local_channel_idx].hiLIM - channels[local_channel_idx].loLIM);

                    1:
                        channels[local_channel_idx].outputValue := TO_REAL(analogValues[local_analog_idx]) / 10.0;

                    2:
                        channels[local_channel_idx].outputValue := TO_REAL(analogValues[local_analog_idx]) / 100.0;
                END_CASE;
            END_IF;
        ELSE
            (* disabled: no writes to retVal or outputValue *)
        END_IF;
    END_FOR;
END_IF;

END_FUNCTION_BLOCK
